// Команды по умолчанию
Command.stIo.xOpenDoor := FALSE;
Command.stIo.xCloseDoor := FALSE;
Command.stIo.xHatchUnLock := FALSE;
Command.stIo.xOpenSafetyDoor := FALSE;
Command.stIo.xCloseSafetyDoor := FALSE;
Command.stIo.xClampChuck := FALSE;
Command.stIo.xUnclampChuck := FALSE;
Command.stIo.xStartCycle := FALSE;
Command.stIo.xReset := xReset OR xResetGlobal;

Command.stRobot.xExecute := FALSE;
Command.stRobot.xStop := FALSE;

// Импульсы ручного управления проходят только через рассчитанные PLC-разрешения.
// Автоматический алгоритм станка в DISABLED не формирует параллельных команд.
IF xHmiOpenSafetyDoor AND xManualSafetyDoorOpenAllowed THEN
	Command.stIo.xOpenSafetyDoor := TRUE;
END_IF;
IF xHmiCloseSafetyDoor AND xManualSafetyDoorCloseAllowed THEN
	Command.stIo.xCloseSafetyDoor := TRUE;
END_IF;
IF xHmiOpenHatch AND xManualHatchOpenAllowed THEN
	xManualHatchOpenDemand := TRUE;
	xManualHatchUnlockDemand := TRUE;
END_IF;
IF xHmiCloseHatch AND xManualHatchCloseAllowed THEN
	Command.stIo.xCloseDoor := TRUE;
	xManualHatchOpenDemand := FALSE;
	xManualHatchUnlockDemand := FALSE;
END_IF;
IF rtHmiUnlockHatch.Q AND xManualHatchUnlockAllowed THEN
	xManualHatchUnlockDemand := TRUE;
END_IF;
IF rtHmiLockHatch.Q AND xManualHatchLockAllowed THEN
	xManualHatchUnlockDemand := FALSE;
	xManualHatchOpenDemand := FALSE;
END_IF;
IF NOT xManualMode THEN
	xManualHatchUnlockDemand := FALSE;
	xManualHatchOpenDemand := FALSE;
END_IF;
IF xHmiOpenChuck AND xManualChuckOpenAllowed THEN
	Command.stIo.xUnclampChuck := TRUE;
END_IF;
IF xHmiCloseChuck AND xManualChuckCloseAllowed THEN
	Command.stIo.xClampChuck := TRUE;
END_IF;
Command.stRobot.eAction := E_ROBOT_ACTION.NONE;
xServiceDoorOpenDemand := FALSE;
xServiceDoorCloseDemand := FALSE;
xServiceHatchUnlockDemand := FALSE;

IF xTestInitialize THEN
	Error.dwErrorActive := DWORD#0;
	Error.dwAlarmActive := DWORD#0;
	uiIndex := UINT#0;
	xDisableRequest := FALSE;
	xOperatorRunningCNC := FALSE;
	xOperatorClosingDoor := FALSE;
	xAutoCycleCommanded := FALSE;
	xCycleMeasureActive := FALSE;
	xCycleMeasureValid := FALSE;
	xRetreatStarted := FALSE;
	xRobotInsideMachine := FALSE;
	xFaultContextCaptured := FALSE;
	xRobotInsideAtFault := FALSE;
	xDoorRobotStopLatched := FALSE;
	xRobotStopRequired := FALSE;
	xRobotDone := FALSE;
	xServiceDoorCloseDemand := FALSE;
	xServiceDoorOpenDemand := FALSE;
	xServiceHatchUnlockDemand := FALSE;
	xManualHatchUnlockDemand := FALSE;
	xManualHatchOpenDemand := FALSE;
	xAutoDoorOpenLatched := FALSE;
	xRobotActionDone := FALSE;
	xRobotCommandStarted := FALSE;
	eGrantedOperation := E_MACHINE_OPERATION.NONE;
	eActualOperation := E_MACHINE_OPERATION.NONE;
	IF (uiTestInitialState = UINT#0) OR NOT xPointsConfigured THEN
		eState := E_MACHINE_STATE.DISABLED;
		ePartType := E_PART_TYPE.UNKNOWN;
	ELSE
		eState := E_MACHINE_STATE.IDLE;
		IF uiTestInitialState = UINT#3 THEN
			ePartType := E_PART_TYPE.DETAIL;
		ELSIF uiTestInitialState = UINT#2 THEN
			ePartType := E_PART_TYPE.PART;
		ELSE
			ePartType := E_PART_TYPE.UNKNOWN;
		END_IF;
	END_IF;
END_IF;

IF stMachineStatus.xChuckClamped AND NOT stMachineStatus.xAlarm THEN
	ePartState := E_PART_STATE.LOADED;
ELSIF stMachineStatus.xChuckUnclamped AND NOT stMachineStatus.xAlarm THEN
	ePartState := E_PART_STATE.EMPTY;
ELSE
	ePartState := E_PART_STATE.UNKNOWN;
END_IF


// // Ручное подтверждение состояния детали
// IF (eState = E_MACHINE_STATE.IDLE)
// AND NOT stMachineStatus.xCycleActive THEN
//     IF rtSetPartLoaded.Q THEN
//         ePartState := E_PART_STATE.LOADED;
//     END_IF;
// 
//     IF rtSetPartEmpty.Q THEN
//         ePartState := E_PART_STATE.EMPTY;
//     END_IF;
// END_IF;

// Автоматическое открытие после окончания обработки
IF rtCycleDone.Q 
	AND NOT stMachineStatus.xAlarm 
	AND NOT stMachineStatus.xCycleActive 
	AND (eState = E_MACHINE_STATE.IDLE) 
	AND NOT xGlobalError THEN
	ePartType := E_PART_TYPE.DETAIL;
    xAutoDoorOpenLatched := TRUE;
END_IF;

IF stMachineStatus.xDoorOpen THEN
    xAutoDoorOpenLatched := FALSE;
END_IF;

eGrantedOperation := E_MACHINE_OPERATION.NONE;

IF (ePartState = E_PART_STATE.EMPTY)
AND (ePartType = E_PART_TYPE.UNKNOWN)
AND stRobotStatus.xBlankAvailable  THEN
    eGrantedOperation := E_MACHINE_OPERATION.LOAD;

ELSIF (ePartState = E_PART_STATE.LOADED)
AND (ePartType = E_PART_TYPE.DETAIL) THEN
    IF stRobotStatus.xBlankAvailable THEN
        eGrantedOperation := E_MACHINE_OPERATION.CHANGE;
    ELSE
        eGrantedOperation := E_MACHINE_OPERATION.UNLOAD;
    END_IF;
ELSIF (ePartState = E_PART_STATE.UNKNOWN) THEN
	eGrantedOperation := E_MACHINE_OPERATION.NONE;
END_IF;

// Включение и отключение блока
IF xDisableRequest
AND ((eState = E_MACHINE_STATE.IDLE)
	OR (eState = E_MACHINE_STATE.OPERATOR_CHOICE_PART)
	OR (eState = E_MACHINE_STATE.OPERATOR_CHOICE_DOOR)
	OR (eState = E_MACHINE_STATE.OPERATOR_CHOICE_RUN)) THEN
    eState := E_MACHINE_STATE.DISABLED;
ELSIF rtEnabledMachine.Q
AND NOT rtDisabledMachine.Q
AND (eState = E_MACHINE_STATE.DISABLED) THEN
	IF NOT stMachineStatus.xAlarm
	AND NOT stMachineStatus.xCycleActive
	AND xSafetyDoorSafe
	AND xPointsConfigured THEN
		IF ePartState = E_PART_STATE.EMPTY THEN
			eState := E_MACHINE_STATE.IDLE;
		ELSIF ePartState = E_PART_STATE.LOADED THEN
			eState := E_MACHINE_STATE.OPERATOR_CHOICE_PART;
		END_IF;
	END_IF;
END_IF;

IF xGlobalError
AND (eState <> E_MACHINE_STATE.DISABLED) THEN
    Error.dwErrorActive := Error.dwErrorActive OR ERR_SAFETY_STOP;
    eState := E_MACHINE_STATE.ERROR;
END_IF;

IF stMachineStatus.xAlarm AND (eState = E_MACHINE_STATE.IDLE) THEN
	Error.dwErrorActive := Error.dwErrorActive OR ERR_MACHINE_IDLE;
    eState := E_MACHINE_STATE.ERROR;
END_IF

IF ((eState = E_MACHINE_STATE.OPERATOR_CHOICE_PART) OR (eState = E_MACHINE_STATE.OPERATOR_CHOICE_DOOR) OR (eState = E_MACHINE_STATE.OPERATOR_CHOICE_RUN))
AND ftChuckClamped.Q THEN
	eState := E_MACHINE_STATE.DISABLED;
END_IF; 

IF (eState = E_MACHINE_STATE.DISABLED) OR (eState = E_MACHINE_STATE.ERROR) THEN
	xOperatorRunningCNC := FALSE;
	xOperatorClosingDoor := FALSE;
	ePartType :=   E_PART_TYPE.UNKNOWN;
END_IF
// Останавливаем робота, если люк закрылся при нахождении робота в станке.
tofErrorDoor(
			PT:= T#100MS,
			IN:=stMachineStatus.xDoorOpen
);

// Ошибка робота в рабочей зоне принадлежит одновременно роботу и станку.
// Для действия захвата сохраняется отдельная диагностическая причина.
IF xRobotInsideMachine
AND stRobotStatus.xError
AND (eState <> E_MACHINE_STATE.ERROR) THEN
	IF eState = E_MACHINE_STATE.ROBOT_ACTION THEN
		Error.dwErrorActive := Error.dwErrorActive OR ERR_ROBOT_ACTION;
	ELSE
		Error.dwErrorActive := Error.dwErrorActive OR ERR_ROBOT_MOTION;
	END_IF;
	eState := E_MACHINE_STATE.ERROR;
END_IF;
						
IF xRobotInsideMachine
AND (
	(rtDoorClosed.Q)
	OR (
		NOT tofErrorDoor.Q
		AND (stRobotStatus.xBusy
			OR (eState = E_MACHINE_STATE.ROBOT_MOVE)
			OR (eState = E_MACHINE_STATE.ROBOT_ACTION))
	)
) THEN
	// Stop должен быть явным даже при гонке статусов: xBusy уже мог успеть
	// сброситься в FB_ROBOT, пока группа ещё принимает команду останова.
	Command.stRobot.xStop := TRUE;
	xDoorRobotStopLatched := TRUE;
	Error.dwErrorActive := Error.dwErrorActive OR ERR_DOOR_ROBOT;
    eState := E_MACHINE_STATE.ERROR;
END_IF

// Открытие операторской двери в любой момент роботного обслуживания
// — первичная авария станка с каскадным ROBOT_STOP.
IF (eActualOperation <> E_MACHINE_OPERATION.NONE)
AND NOT xManualMode
AND NOT xSafetyDoorSafe
AND (eState <> E_MACHINE_STATE.ERROR) THEN
	Command.stRobot.xStop := stRobotStatus.xBusy;
	Error.dwErrorActive := Error.dwErrorActive OR ERR_SAFETY_DOOR_OPEN;
	eState := E_MACHINE_STATE.ERROR;
END_IF;

// Старый рецепт и удерживаемые запросы не возобновляются после ручного I/O.
// Состояние патрона будет повторно определено при отдельном включении станка.
IF xIoManual THEN
	uiIndex := UINT#0;
	eActualOperation := E_MACHINE_OPERATION.NONE;
	eGrantedOperation := E_MACHINE_OPERATION.NONE;
	xRobotDone := FALSE;
	xRobotCommandStarted := FALSE;
	xManualHatchUnlockDemand := FALSE;
	xManualHatchOpenDemand := FALSE;
	xAutoDoorOpenLatched := FALSE;
	xOperatorRunningCNC := FALSE;
	xOperatorClosingDoor := FALSE;
	IF eState <> E_MACHINE_STATE.ERROR THEN
		eState := E_MACHINE_STATE.DISABLED;
	END_IF;
END_IF;

CASE eState OF
	E_MACHINE_STATE.DISABLED:
		xDisableRequest := FALSE;
		IF NOT stMachineStatus.xCycleActive THEN
			xAutoCycleCommanded := FALSE;
		END_IF;
		
	E_MACHINE_STATE.OPERATOR_CHOICE_PART:
		IF rtSetDetailLoaded.Q AND NOT stMachineStatus.xAlarm THEN
			eState := E_MACHINE_STATE.IDLE;
			ePartType := E_PART_TYPE.DETAIL;
		ELSIF rtSetBlankLoaded.Q AND NOT stMachineStatus.xAlarm THEN
			ePartType := E_PART_TYPE.PART;
			IF stMachineStatus.xDoorClosed THEN
				eState := E_MACHINE_STATE.OPERATOR_CHOICE_RUN;
			ELSE
				eState := E_MACHINE_STATE.OPERATOR_CHOICE_DOOR;
			END_IF;
		ELSIF stMachineStatus.xAlarm THEN
			Error.dwErrorActive := Error.dwErrorActive OR ERR_MACHINE_ALARM;
    		eState := E_MACHINE_STATE.ERROR;
		END_IF;
		
	E_MACHINE_STATE.OPERATOR_CHOICE_DOOR:
		// При уже закрытой двери шаг подтверждения закрытия не нужен:
		// автомат сразу переходит к вопросу о запуске обработки.
		IF stMachineStatus.xAlarm THEN
			Error.dwErrorActive := Error.dwErrorActive OR ERR_MACHINE_ALARM;
    		eState := E_MACHINE_STATE.ERROR;
		ELSIF xHmiRejectDoor THEN
			eState := E_MACHINE_STATE.DISABLED;
		ELSIF stMachineStatus.xDoorClosed THEN
			eState := E_MACHINE_STATE.OPERATOR_CHOICE_RUN;
		ELSIF xHmiAcceptDoor THEN
			xOperatorClosingDoor := TRUE;
			eState := E_MACHINE_STATE.DOOR_CLOSE;
		END_IF;
		
	E_MACHINE_STATE.OPERATOR_CHOICE_RUN:
		IF xHmiAcceptRunCNC AND NOT stMachineStatus.xAlarm THEN
			xOperatorRunningCNC := TRUE; 
			eState := E_MACHINE_STATE.CYCLE_START;
		ELSIF xHmiRejectRunCNC AND NOT stMachineStatus.xAlarm THEN
			eState := E_MACHINE_STATE.DISABLED;
		ELSIF stMachineStatus.xAlarm THEN
			Error.dwErrorActive := Error.dwErrorActive OR ERR_MACHINE_ALARM;
    		eState := E_MACHINE_STATE.ERROR;
		END_IF; 	
		
	E_MACHINE_STATE.IDLE:
		uiIndex := 0;
		xRobotDone := FALSE;
		IF xExecute THEN
			IF (stRobotStatus.eCurrentPoint = stPoints.eAbove)
			AND ePartState <> E_PART_STATE.UNKNOWN
			AND NOT stMachineStatus.xAlarm
			AND NOT stMachineStatus.xCycleActive
			AND xSafetyDoorSafe
    		AND NOT stRobotStatus.xBusy 
			AND NOT stRobotStatus.xError
			AND NOT xGlobalError THEN
				eActualOperation := eGrantedOperation;
				eState := E_MACHINE_STATE.CHOSE;
			ELSIF ePartState = E_PART_STATE.UNKNOWN THEN
				Error.dwErrorActive := Error.dwErrorActive OR ERR_UNKNOWN_DETAIL;
				eState := E_MACHINE_STATE.ERROR ;
			END_IF
		END_IF
		
	E_MACHINE_STATE.CHOSE:
		CASE eActualOperation OF 
			E_MACHINE_OPERATION.CHANGE:
				stRecipe := stChangeRecipe;
				eState := E_MACHINE_STATE.READ;
			E_MACHINE_OPERATION.LOAD:
				stRecipe := stLoadRecipe;
				eState := E_MACHINE_STATE.READ;
			E_MACHINE_OPERATION.UNLOAD:
				stRecipe := stUnloadRecipe;
				eState := E_MACHINE_STATE.READ;
		ELSE
			Error.dwErrorActive := Error.dwErrorActive OR ERR_WRONG_OPERATION ;
			eState := E_MACHINE_STATE.ERROR;
		END_CASE
		
	E_MACHINE_STATE.READ:
		CASE stRecipe[uiIndex].eCommand OF
			E_MACHINE_STATE.ROBOT_MOVE:
				xRobotCommandStarted := FALSE;
				eState := E_MACHINE_STATE.ROBOT_MOVE;
				
			E_MACHINE_STATE.ROBOT_ACTION:
				xRobotCommandStarted := FALSE;
				eState := E_MACHINE_STATE.ROBOT_ACTION;
				
			E_MACHINE_STATE.DOOR_OPEN:
				eState := E_MACHINE_STATE.DOOR_OPEN;
				
			E_MACHINE_STATE.DOOR_CLOSE:
				eState := E_MACHINE_STATE.DOOR_CLOSE;
				
			E_MACHINE_STATE.CHUCK_OPEN:
				eState := E_MACHINE_STATE.CHUCK_OPEN;
				
			E_MACHINE_STATE.CHUCK_CLOSE:
				eState := E_MACHINE_STATE.CHUCK_CLOSE;
				
			E_MACHINE_STATE.CYCLE_START:
				eState := E_MACHINE_STATE.CYCLE_START;
				
			E_MACHINE_STATE.DONE:
				eState := E_MACHINE_STATE.DONE;
				
		ELSE
			Error.dwErrorActive := Error.dwErrorActive OR ERR_WRONG_COMMAND;
			eState := E_MACHINE_STATE.ERROR;
		END_CASE
	
	E_MACHINE_STATE.NEXT:
			uiIndex := uiIndex + 1;
			IF uiIndex > 40 THEN
				Error.dwErrorActive := Error.dwErrorActive OR ERR_INDEX;
				eState := E_MACHINE_STATE.ERROR;
			ELSE
				eState := E_MACHINE_STATE.READ;
			END_IF;
	
	E_MACHINE_STATE.ROBOT_MOVE:
		Command.stRobot.xExecute  := TRUE;
		Command.stRobot.eAction   := E_ROBOT_ACTION.MOVE_TO_POINT;
		xRetreatStarted          := stRecipe[uiIndex].xRetreatStarted;
		IF stRecipe[uiIndex].stPoint = E_MACHINE_POINTS.ABOVE  THEN
			Command.stRobot.eSetPoint := stPoints.eAbove;
		ELSIF stRecipe[uiIndex].stPoint = E_MACHINE_POINTS.CHUCK THEN
			Command.stRobot.eSetPoint := stPoints.eChuck;
		ELSIF stRecipe[uiIndex].stPoint = E_MACHINE_POINTS.CHUCK_APPROACH THEN
			Command.stRobot.eSetPoint := stPoints.eChuckApproach;
		ELSIF stRecipe[uiIndex].stPoint = E_MACHINE_POINTS.INSIDE THEN
			Command.stRobot.eSetPoint := stPoints.eInside;
		END_IF
		IF stRobotStatus.xBusy THEN
			xRobotCommandStarted := TRUE;
		END_IF;

		IF stRobotStatus.xError THEN
			Error.dwErrorActive := Error.dwErrorActive OR ERR_ROBOT_MOTION;
			eState := E_MACHINE_STATE.ERROR ;
			
		ELSIF stMachineStatus.xAlarm THEN
			Command.stRobot.xStop := stRobotStatus.xBusy;
			Error.dwErrorActive := Error.dwErrorActive OR ERR_MACHINE_ALARM;
			eState := E_MACHINE_STATE.ERROR ;
			
		ELSIF xRobotCommandStarted AND stRobotStatus.xDone THEN
        	eState := E_MACHINE_STATE.RELEASE_ROBOT_ACTION;

		ELSIF tonRobotMoveTimeout.Q THEN
			Command.stRobot.xStop := stRobotStatus.xBusy;
			Error.dwErrorActive := Error.dwErrorActive OR ERR_TIMEOUT_ROBOT_MOVE;
			eState := E_MACHINE_STATE.ERROR;
			
    	END_IF;
	
	E_MACHINE_STATE.ROBOT_ACTION:
		xRobotActionDone := FALSE;

		CASE stRecipe[uiIndex].eRobotAction OF
			E_ROBOT_ACTION.UNCLAMP_1:
				xRobotActionDone := stRobotStatus.xGripper1Open;
			E_ROBOT_ACTION.CLAMP_1:
				xRobotActionDone := stRobotStatus.xGripper1Closed;
			E_ROBOT_ACTION.UNCLAMP_2:
				xRobotActionDone := stRobotStatus.xGripper2Open;
			E_ROBOT_ACTION.CLAMP_2:
				xRobotActionDone := stRobotStatus.xGripper2Closed;
			E_ROBOT_ACTION.ROTATE_TO_BLANK:
				xRobotActionDone := stRobotStatus.xRotatedToBlank;
			E_ROBOT_ACTION.ROTATE_TO_DETAIL:
				xRobotActionDone := stRobotStatus.xRotatedToDetail;
		END_CASE;
		IF xRobotActionDone THEN
			eState := E_MACHINE_STATE.NEXT;
		ELSE
			Command.stRobot.xExecute := TRUE;
			Command.stRobot.eAction := stRecipe[uiIndex].eRobotAction;
		END_IF;
		IF stRobotStatus.xBusy THEN
			xRobotCommandStarted := TRUE;
		END_IF;
		
		IF (eState = E_MACHINE_STATE.ROBOT_ACTION)
		AND stMachineStatus.xAlarm THEN
			Command.stRobot.xStop := stRobotStatus.xBusy;
			Error.dwErrorActive := Error.dwErrorActive OR ERR_MACHINE_ALARM;
			eState := E_MACHINE_STATE.ERROR ;
	
		ELSIF (eState = E_MACHINE_STATE.ROBOT_ACTION)
		AND stRobotStatus.xError THEN
			Error.dwErrorActive := Error.dwErrorActive OR ERR_ROBOT_ACTION;
			eState := E_MACHINE_STATE.ERROR ;

		ELSIF (eState = E_MACHINE_STATE.ROBOT_ACTION)
		AND tonRobotActionTimeout.Q THEN
			Command.stRobot.xStop := stRobotStatus.xBusy;
			Error.dwErrorActive := Error.dwErrorActive OR ERR_TIMEOUT_ROBOT_ACTION;
			eState := E_MACHINE_STATE.ERROR;
			
		ELSIF (eState = E_MACHINE_STATE.ROBOT_ACTION)
		AND xRobotCommandStarted
		AND stRobotStatus.xDone THEN
        	eState := E_MACHINE_STATE.RELEASE_ROBOT_ACTION;
    	END_IF;
		
	E_MACHINE_STATE.RELEASE_ROBOT_ACTION:
		IF NOT stRobotStatus.xBusy
    	AND NOT stRobotStatus.xDone
		AND NOT stRobotStatus.xError THEN
			xRobotDone := stRecipe[uiIndex].xRobotDone;
        	eState := E_MACHINE_STATE.NEXT;
			
		ELSIF stRobotStatus.xError AND  stRecipe[uiIndex].eRobotAction = E_ROBOT_ACTION.MOVE_TO_POINT THEN
			Error.dwErrorActive := Error.dwErrorActive OR ERR_ROBOT_MOTION;
			eState := E_MACHINE_STATE.ERROR;
			
		ELSIF stRobotStatus.xError THEN
			Error.dwErrorActive := Error.dwErrorActive OR ERR_ROBOT_ACTION;
			eState := E_MACHINE_STATE.ERROR;

		ELSIF tonRobotReleaseTimeout.Q THEN
			Command.stRobot.xStop := stRobotStatus.xBusy;
			Error.dwErrorActive := Error.dwErrorActive OR ERR_TIMEOUT_ROBOT_RELEASE;
			eState := E_MACHINE_STATE.ERROR;
    	END_IF;
		
	E_MACHINE_STATE.DOOR_OPEN:
		xServiceDoorOpenDemand := TRUE;
		// Сначала снимаем замок, затем открываем роботный люк.
		IF stMachineStatus.xHatchLocked THEN
			xServiceHatchUnlockDemand := TRUE;
		END_IF;

	    IF stMachineStatus.xDoorOpen
		AND NOT stMachineStatus.xHatchLocked
		AND NOT stMachineStatus.xAlarm THEN
			xServiceDoorOpenDemand := FALSE;
			xServiceHatchUnlockDemand := FALSE;
         	eState := E_MACHINE_STATE.NEXT;
		ELSIF stMachineStatus.xAlarm THEN
			Error.dwErrorActive := Error.dwErrorActive OR ERR_DOOR_OPEN;
			eState := E_MACHINE_STATE.ERROR;
		ELSIF tonDoorOpenTimeout.Q THEN
			xServiceDoorOpenDemand := FALSE;
			Error.dwErrorActive := Error.dwErrorActive OR ERR_TIMEOUT_DOOR_OPEN;
			eState := E_MACHINE_STATE.ERROR;
    	END_IF;
	
	E_MACHINE_STATE.DOOR_CLOSE: 
		// После сервисной операции безопасность подтверждает защёлка xRobotDone:
		// рецепт уже довёл робот до ABOVE и освободил его для следующего маршрута.
		// Общий xBusy больше не блокирует дверь: робот может двигаться к другому узлу.
		IF xRobotInsideMachine
		OR (NOT xOperatorClosingDoor AND NOT xRobotDone) THEN
			Command.stRobot.xStop := xRobotInsideMachine AND stRobotStatus.xBusy;
			xDoorRobotStopLatched := TRUE;
			Error.dwErrorActive := Error.dwErrorActive OR ERR_DOOR_ROBOT;
			eState := E_MACHINE_STATE.ERROR;
		ELSE
			xServiceDoorCloseDemand := TRUE;
			// Замок удерживается открытым до подтверждения закрытой двери.
			IF NOT stMachineStatus.xDoorClosed THEN
				xServiceHatchUnlockDemand := TRUE;
			END_IF;
		END_IF;

		IF stMachineStatus.xDoorClosed THEN
			xServiceHatchUnlockDemand := FALSE;
		END_IF;
		IF (eState = E_MACHINE_STATE.DOOR_CLOSE)
		AND stMachineStatus.xDoorClosed
		AND stMachineStatus.xHatchLocked
		AND NOT stMachineStatus.xAlarm THEN
			xServiceDoorCloseDemand := FALSE;
			IF NOT xOperatorClosingDoor THEN
				eState := E_MACHINE_STATE.NEXT;
			ELSIF xOperatorClosingDoor THEN
				eState := E_MACHINE_STATE.OPERATOR_CHOICE_RUN;
				xOperatorClosingDoor := FALSE;
			END_IF;
		ELSIF stMachineStatus.xAlarm THEN
			Error.dwErrorActive := Error.dwErrorActive OR ERR_DOOR_CLOSE;
			eState := E_MACHINE_STATE.ERROR;
		ELSIF (eState = E_MACHINE_STATE.DOOR_CLOSE)
		AND tonDoorCloseTimeout.Q THEN
			xServiceDoorCloseDemand := FALSE;
			Error.dwErrorActive := Error.dwErrorActive OR ERR_TIMEOUT_DOOR_CLOSE;
			eState := E_MACHINE_STATE.ERROR;
    	END_IF;
		
	E_MACHINE_STATE.CHUCK_OPEN: 
		Command.stIo.xUnclampChuck := TRUE;

    	IF stMachineStatus.xChuckUnclamped 
		AND NOT stMachineStatus.xAlarm THEN
			Command.stIo.xUnclampChuck := FALSE;
			ePartType := E_PART_TYPE.UNKNOWN;
       		eState := E_MACHINE_STATE.NEXT;
		ELSIF stMachineStatus.xAlarm THEN
			Command.stIo.xUnclampChuck := FALSE;
			Error.dwErrorActive := Error.dwErrorActive OR ERR_CHUCK_OPEN;
			eState := E_MACHINE_STATE.ERROR;
		ELSIF tonChuckOpenTimeout.Q THEN
			Command.stIo.xUnclampChuck := FALSE;
			Error.dwErrorActive := Error.dwErrorActive OR ERR_TIMEOUT_CHUCK_OPEN;
			eState := E_MACHINE_STATE.ERROR;
    	END_IF;
		
	
	E_MACHINE_STATE.CHUCK_CLOSE: 
		Command.stIo.xClampChuck := TRUE;

    	IF stMachineStatus.xChuckClamped 
		AND NOT stMachineStatus.xAlarm THEN
			Command.stIo.xClampChuck := FALSE;
			ePartType := E_PART_TYPE.PART;
       		eState := E_MACHINE_STATE.NEXT;
		ELSIF stMachineStatus.xAlarm THEN
			Command.stIo.xClampChuck := FALSE;
			Error.dwErrorActive := Error.dwErrorActive OR ERR_CHUCK_CLOSE;
			eState := E_MACHINE_STATE.ERROR;
		ELSIF tonChuckCloseTimeout.Q THEN
			Command.stIo.xClampChuck := FALSE;
			Error.dwErrorActive := Error.dwErrorActive OR ERR_TIMEOUT_CHUCK_CLOSE;
			eState := E_MACHINE_STATE.ERROR;
    	END_IF;
		
	E_MACHINE_STATE.CYCLE_START:
		IF stMachineStatus.xChuckClamped
    	AND stMachineStatus.xDoorClosed THEN
			Command.stIo.xStartCycle := TRUE;
			xAutoCycleCommanded := TRUE;
		END_IF;
		
        IF stMachineStatus.xCycleActive
		AND NOT stMachineStatus.xAlarm THEN
			Command.stIo.xStartCycle := FALSE;
			IF NOT xOperatorRunningCNC THEN
            	eState := E_MACHINE_STATE.NEXT;
			ELSIF xOperatorRunningCNC THEN
				xOperatorRunningCNC := FALSE;
				eState := E_MACHINE_STATE.IDLE;
			END_IF;
		ELSIF stMachineStatus.xAlarm THEN
			Command.stIo.xStartCycle := FALSE;
			Error.dwErrorActive := Error.dwErrorActive OR ERR_CYCLE_START;
			eState := E_MACHINE_STATE.ERROR;
		ELSIF tonCycleStartTimeout.Q THEN
			Command.stIo.xStartCycle := FALSE;
			xAutoCycleCommanded := FALSE;
			Error.dwErrorActive := Error.dwErrorActive OR ERR_TIMEOUT_CYCLE_START;
			eState := E_MACHINE_STATE.ERROR;
        END_IF;
	
	E_MACHINE_STATE.DONE:
		CASE eActualOperation OF 
			E_MACHINE_OPERATION.CHANGE, E_MACHINE_OPERATION.LOAD:
				eActualOperation := E_MACHINE_OPERATION.NONE;
				ePartState := E_PART_STATE.LOADED;						
			E_MACHINE_OPERATION.UNLOAD:
				eActualOperation := E_MACHINE_OPERATION.NONE;
				ePartState := E_PART_STATE.EMPTY;
		END_CASE
		
		IF NOT xExecute THEN
			xRobotDone := FALSE;	
			eState := E_MACHINE_STATE.IDLE;
		END_IF
		
    E_MACHINE_STATE.ERROR:
		uiIndex := 0;
		eActualOperation := E_MACHINE_OPERATION.NONE;
		eGrantedOperation := E_MACHINE_OPERATION.NONE;
		IF NOT stMachineStatus.xCycleActive THEN
			xAutoCycleCommanded := FALSE;
		END_IF;

		IF (xReset OR xResetGlobal)
		AND NOT xIoManual
		AND NOT xGlobalError
		AND NOT xExecute
		AND NOT stMachineStatus.xAlarm
		AND xSafetyDoorSafe
		AND xDoorRobotRecoveryReady
		AND xRobotResetDependencyReady THEN
			Error.dwErrorLast := Error.dwErrorActive;
			Error.dwErrorActive := DWORD#0;
			xManualHatchUnlockDemand := FALSE;
			xManualHatchOpenDemand := FALSE;
        	eState := E_MACHINE_STATE.DISABLED;
    	END_IF;
END_CASE;

// Таймаут одинаково контролирует автоматическое и ручное снятие замка.
// После отказа удерживаемый запрос снимается, чтобы сброс не запустил его
// повторно без нового явного действия оператора.
IF tonHatchUnlockTimeout.Q
AND (eState <> E_MACHINE_STATE.ERROR) THEN
	xServiceHatchUnlockDemand := FALSE;
	xManualHatchUnlockDemand := FALSE;
	xManualHatchOpenDemand := FALSE;
	Error.dwErrorActive := Error.dwErrorActive OR ERR_TIMEOUT_HATCH_UNLOCK;
	eState := E_MACHINE_STATE.ERROR;
END_IF;

// Причина остаётся в своём CASE, а единая реакция рассчитывается один раз.
// Контекст защёлкивается до сброса, поэтому смена состояния робота его не теряет.
IF (eState = E_MACHINE_STATE.ERROR) AND NOT xFaultContextCaptured THEN
	xRobotInsideAtFault := xRobotInsideMachine;
	xFaultContextCaptured := TRUE;
ELSIF eState <> E_MACHINE_STATE.ERROR THEN
	xRobotInsideAtFault := FALSE;
	xFaultContextCaptured := FALSE;
END_IF;

xRobotStopRequired := NOT xGlobalError
	AND (
		((Error.dwErrorActive
			AND (MASK_ALWAYS_ROBOT_STOP AND NOT ERR_DOOR_ROBOT)) <> DWORD#0)
		OR (((Error.dwErrorActive AND ERR_DOOR_ROBOT) <> DWORD#0)
			AND NOT xDoorRobotRecoveryReady)
		OR xDoorRobotStopLatched
		OR (((Error.dwErrorActive
			AND (MASK_EQUIPMENT_ERROR AND NOT ERR_DOOR_ROBOT)) <> DWORD#0)
			AND xRobotInsideAtFault)
	);

// Stop нужен только выполняемому действию. Стоящий в станке робот получает
// зависимую ошибку через FB_ROBOT, но бессмысленная команда Stop не выдаётся.
IF (eState = E_MACHINE_STATE.ERROR)
AND xRobotStopRequired
AND (stRobotStatus.xBusy OR xRobotMotionBusy) THEN
	Command.stRobot.xStop := TRUE;
END_IF;

// После подтверждённого открытия люка и полной остановки можно отпустить
// защёлку зависимого Stop; до этого новый цикл не должен стартовать.
IF xDoorRobotStopLatched
AND NOT xRobotMotionBusy
AND xDoorRobotRecoveryReady THEN
	xDoorRobotStopLatched := FALSE;
END_IF;

IF ((eState <> E_MACHINE_STATE.ERROR) OR xManualHatchRecoveryOpenAllowed)
AND NOT xGlobalError AND NOT xIoManual THEN
	Command.stIo.xHatchUnLock := xManualHatchUnlockDemand OR xServiceHatchUnlockDemand;
	IF xManualHatchOpenDemand
	AND NOT stMachineStatus.xHatchLocked
	AND NOT stMachineStatus.xDoorOpen
	AND NOT stMachineStatus.xCycleActive
	AND NOT stMachineStatus.xAlarm THEN
		Command.stIo.xOpenDoor := TRUE;
	END_IF;
    IF (eState <> E_MACHINE_STATE.ERROR) AND xServiceDoorCloseDemand 
	AND NOT (xAutoDoorOpenLatched OR xServiceDoorOpenDemand)
	AND NOT xRobotInsideMachine
	AND (xOperatorClosingDoor OR xRobotDone)
	AND NOT stMachineStatus.xAlarm THEN
        Command.stIo.xCloseDoor := TRUE;

    ELSIF (eState <> E_MACHINE_STATE.ERROR) AND (xAutoDoorOpenLatched OR xServiceDoorOpenDemand)
	AND NOT xServiceDoorCloseDemand
	AND NOT stMachineStatus.xHatchLocked
    AND NOT stMachineStatus.xCycleActive
    AND NOT stMachineStatus.xAlarm THEN
        Command.stIo.xOpenDoor := TRUE;
    END_IF;
END_IF;

// Замок нельзя открывать во время обработки выбранного для автоматической
// линии станка. Срабатывание формируется самим PLC по фактической команде.
IF xAutomaticUseEnabled
AND stMachineStatus.xCycleActive
AND NOT stMachineStatus.xHatchLocked THEN
	Command.stIo.xHatchUnLock := FALSE;
	Error.dwErrorActive := Error.dwErrorActive OR ERR_HATCH_UNLOCK_PROCESSING;
	eState := E_MACHINE_STATE.ERROR;
END_IF;

Status.xCanAcceptService := (eState = E_MACHINE_STATE.IDLE)
			AND ePartState <> E_PART_STATE.UNKNOWN
			AND NOT stMachineStatus.xAlarm
			AND NOT stMachineStatus.xCycleActive
			AND xSafetyDoorSafe
			AND NOT xGlobalError;

// В состоянии ERROR станок уже остановлен и не считается включённым.
// Это позволяет HMI показать команду «Включить станок», но оставить её
// недоступной до устранения причины и сброса ошибки.
Status.xEnabled := (eState <> E_MACHINE_STATE.DISABLED)
	AND (eState <> E_MACHINE_STATE.ERROR);
Status.xDisablePending := xDisableRequest AND Status.xEnabled;
Status.xPowerAllowed := (eState <> E_MACHINE_STATE.ERROR)
	AND (xDisableRequest
		OR (eState <> E_MACHINE_STATE.DISABLED)
		OR ((eState = E_MACHINE_STATE.DISABLED)
			AND xPointsConfigured
			AND NOT stMachineStatus.xAlarm
			AND NOT stMachineStatus.xCycleActive
			AND xSafetyDoorSafe
			AND (ePartState <> E_PART_STATE.UNKNOWN)));
Status.xResetAllowed := (eState = E_MACHINE_STATE.ERROR)
	AND NOT xIoManual
	AND (Error.dwErrorActive <> DWORD#0)
	AND NOT stMachineStatus.xAlarm
	AND xSafetyDoorSafe
	AND NOT xGlobalError
	AND NOT xExecute
	AND (((Error.dwErrorActive AND ERR_DOOR_ROBOT) = DWORD#0)
		OR xDoorRobotRecoveryReady)
	AND xRobotResetDependencyReady;
Status.xManualControlAllowed := xManualControlAllowed;
Status.xManualSafetyDoorControlEnabled := xSafetyDoorControlEnabled;
Status.xManualSafetyDoorOpenAllowed := xManualSafetyDoorOpenAllowed;
Status.xManualSafetyDoorCloseAllowed := xManualSafetyDoorCloseAllowed;
Status.xManualHatchOpenAllowed := xManualHatchOpenAllowed;
Status.xManualHatchCloseAllowed := xManualHatchCloseAllowed;
Status.xManualHatchUnlockAllowed := xManualHatchUnlockAllowed;
Status.xManualHatchLockAllowed := xManualHatchLockAllowed;
Status.xManualChuckOpenAllowed := xManualChuckOpenAllowed;
Status.xManualChuckCloseAllowed := xManualChuckCloseAllowed;
Status.xProcessing := stMachineStatus.xCycleActive;
Status.xPartReady := stMachineStatus.xCycleDone;
Status.xServiceRequired := (eGrantedOperation <> E_MACHINE_OPERATION.NONE)
	AND (eState = E_MACHINE_STATE.IDLE);
Status.xRobotReleased := xRobotDone;
Status.xDone := (eState = E_MACHINE_STATE.DONE);
Status.xBusy :=  (eState <> E_MACHINE_STATE.IDLE)
				AND (eState <> E_MACHINE_STATE.DISABLED)
				AND (eState <> E_MACHINE_STATE.ERROR)
				AND (eState <> E_MACHINE_STATE.DONE)
				AND (eState <> E_MACHINE_STATE.OPERATOR_CHOICE_PART)
				AND (eState <> E_MACHINE_STATE.OPERATOR_CHOICE_RUN)
				AND (eState <> E_MACHINE_STATE.OPERATOR_CHOICE_DOOR)
				AND NOT ((eState = E_MACHINE_STATE.CYCLE_START) AND xOperatorRunningCNC)
				AND NOT ((eState = E_MACHINE_STATE.DOOR_CLOSE) AND xOperatorClosingDoor);
Status.xError := (eState = E_MACHINE_STATE.ERROR);
Status.xCriticalError := xRobotStopRequired;
Status.xAlarmError    := (Error.dwErrorActive AND MASK_EQUIPMENT_ERROR) <> DWORD#0;
Status.xExternalError := (Error.dwErrorActive AND MASK_EXTERNAL_ERROR) <> DWORD#0;
Status.xServiceRejected := (Error.dwErrorActive
	AND (ERR_DOOR_OPEN OR ERR_TIMEOUT_DOOR_OPEN)) <> DWORD#0
	AND ((Error.dwErrorActive
		AND NOT (ERR_DOOR_OPEN OR ERR_TIMEOUT_DOOR_OPEN)) = DWORD#0);
Error.dwAlarmActive := Error.dwErrorActive;
Status.xDoorOpen := stMachineStatus.xDoorOpen;
Status.xAlarm := stMachineStatus.xAlarm;
Status.eRecommendedOperation := eGrantedOperation;
Status.ePartState := ePartState;
Status.ePartType := ePartType;
Status.eAbovePoint := stPoints.eAbove;
Status.tCycleExpected := tExpectedCycle;
Status.tCycleElapsed := tonCycleMeasure.ET;
Status.tMeasuredCycle := tMeasuredCycle;
Status.xCycleTimeValid := tExpectedCycle > T#0S;
Status.xMeasuredTimeValid := xMeasuredTimeValid;
Status.xCycleOvertime := FALSE;
Status.tRemaining := T#0S;

IF stMachineStatus.xCycleActive
AND Status.xCycleTimeValid THEN
	IF Status.tCycleElapsed < Status.tCycleExpected THEN
		Status.tRemaining := Status.tCycleExpected - Status.tCycleElapsed;
	ELSE
		Status.xCycleOvertime := TRUE;
	END_IF;
END_IF;

Diag.eState := eState;
Diag.eGrantedOperation := eGrantedOperation;
Diag.eActualOperation := eActualOperation;

IF Error.dwErrorActive <> DWORD#0 THEN
	Error.dwErrorLast := Error.dwErrorActive;
END_IF;

Error.stErrorActive := UpdateErrorView(dwError := Error.dwErrorActive);
Error.stErrorLast := UpdateErrorView(dwError := Error.dwErrorLast);

METHOD UpdateErrorView : ST_MACHINE_ERROR
VAR_INPUT
	dwError : DWORD; // Битовая маска для расшифровки
END_VAR
VAR
	stError : ST_MACHINE_ERROR; // Представление ошибок отдельными флагами
END_VAR
stError.WRONG_OPERATION := (dwError AND ERR_WRONG_OPERATION) <> DWORD#0;
stError.WRONG_COMMAND := (dwError AND ERR_WRONG_COMMAND) <> DWORD#0;
stError.ROBOT_MOTION := (dwError AND ERR_ROBOT_MOTION) <> DWORD#0;
stError.ROBOT_ACTION := (dwError AND ERR_ROBOT_ACTION) <> DWORD#0;
stError.DOOR_OPEN := (dwError AND ERR_DOOR_OPEN) <> DWORD#0;
stError.DOOR_CLOSE := (dwError AND ERR_DOOR_CLOSE) <> DWORD#0;
stError.CHUCK_OPEN := (dwError AND ERR_CHUCK_OPEN) <> DWORD#0;
stError.CHUCK_CLOSE := (dwError AND ERR_CHUCK_CLOSE) <> DWORD#0;
stError.CYCLE_START := (dwError AND ERR_CYCLE_START) <> DWORD#0;
stError.SAFETY_STOP := (dwError AND ERR_SAFETY_STOP) <> DWORD#0;
stError.UNKNOWN_DETAIL := (dwError AND ERR_UNKNOWN_DETAIL) <> DWORD#0;
stError.MACHINE_ALARM := (dwError AND ERR_MACHINE_ALARM) <> DWORD#0;
stError.INDEX_ERROR := (dwError AND ERR_INDEX) <> DWORD#0;
stError.DOOR_ROBOT := (dwError AND ERR_DOOR_ROBOT) <> DWORD#0;
stError.MACHINE_IDLE := (dwError AND ERR_MACHINE_IDLE) <> DWORD#0;
stError.TIMEOUT_ROBOT_MOVE := (dwError AND ERR_TIMEOUT_ROBOT_MOVE) <> DWORD#0;
stError.TIMEOUT_ROBOT_ACTION := (dwError AND ERR_TIMEOUT_ROBOT_ACTION) <> DWORD#0;
stError.TIMEOUT_ROBOT_RELEASE := (dwError AND ERR_TIMEOUT_ROBOT_RELEASE) <> DWORD#0;
stError.TIMEOUT_DOOR_OPEN := (dwError AND ERR_TIMEOUT_DOOR_OPEN) <> DWORD#0;
stError.TIMEOUT_DOOR_CLOSE := (dwError AND ERR_TIMEOUT_DOOR_CLOSE) <> DWORD#0;
stError.TIMEOUT_HATCH_UNLOCK := (dwError AND ERR_TIMEOUT_HATCH_UNLOCK) <> DWORD#0;
stError.TIMEOUT_CHUCK_OPEN := (dwError AND ERR_TIMEOUT_CHUCK_OPEN) <> DWORD#0;
stError.TIMEOUT_CHUCK_CLOSE := (dwError AND ERR_TIMEOUT_CHUCK_CLOSE) <> DWORD#0;
stError.TIMEOUT_CYCLE_START := (dwError AND ERR_TIMEOUT_CYCLE_START) <> DWORD#0;
stError.SAFETY_DOOR_OPEN := (dwError AND ERR_SAFETY_DOOR_OPEN) <> DWORD#0;
stError.HATCH_UNLOCK_PROCESSING := (dwError AND ERR_HATCH_UNLOCK_PROCESSING) <> DWORD#0;

UpdateErrorView := stError;
END_METHOD

END_FUNCTION_BLOCK

// Device/Application/FB/FB_ROBOT
FUNCTION_BLOCK FB_ROBOT
VAR_INPUT
	xUsePhysicalGripperFeedback : BOOL;
	xPhysicalGripperIoReady : BOOL;
	stPhysicalGripperFeedback : ST_GRIPPER_STATUS;
	tPhysicalGripperActionTimeout : TIME := T#10S;
	axMagazineExchangeInProgress : ARRAY [1..2] OF BOOL; // Блокировка адресуется только к меняемому магазину
	xTestInitialize : BOOL;
	auiTestGripperContent : ARRAY [1..2] OF UINT;
	auiTestGripperType : ARRAY [1..2] OF UINT;
	uiTestOrientation : UINT;
	xExternalCommandInhibit : BOOL; // Программный экстренный останов запрещает следующую внешнюю команду
	xSimulationAccelerationEnable : BOOL; // Разрешить ускорение виртуальных таймеров только в симуляции
	uiSimulationTimeFactor : UINT := 1; // Коэффициент виртуального времени 1..100

	stMachine_1_Command : ST_ROBOT_COMMAND; // Команда роботу от первого станка
	stMachine_2_Command : ST_ROBOT_COMMAND; // Команда роботу от второго станка
	stMachine_3_Command : ST_ROBOT_COMMAND; // Команда роботу от третьего станка
	stMagazineCommand   : ST_ROBOT_COMMAND; // Команда роботу от магазина
	stCellCommand       : ST_ROBOT_COMMAND; // Команда позиционирования от менеджера ячейки
	uiBlankPayloadType  : UINT; // Тип заготовки из состояния цикла
	uiDetailPayloadType : UINT; // Тип готовой детали из состояния цикла
	stHmiCommand        : ST_ROBOT_COMMAND; // Ручная команда роботу с HMI
	xReset              : BOOL; // Сброс ошибок робота
    xMode               : BOOL; // Режим робота: TRUE — Modbus, FALSE — SoftMotion
	xManual      		: BOOL; // 1 - ручной режим работы, 0 - автоматический режим работы
	xGlobalError        : BOOL; // Глобальная ошибка ячейки
	xEquipmentStopRequired : BOOL; // Владелец оборудования требует зависимую ошибку робота
	xModbusBusy         : BOOL; // Внешний робот выполняет команду
	xModbusDone         : BOOL; // Внешний робот завершил команду
	xModbusError        : BOOL; // Ошибка обмена или внешнего робота
	stModbusStatus      : ST_ROBOT_MODBUS_STATUS; // Декодированная обратная связь SC-500
	xHmiDrivesEnable    : BOOL; // Исходный запрос HMI на включение приводов
	xHmiDrivesDisable   : BOOL; // Исходный запрос HMI на отключение приводов
	xHmiStop            : BOOL; // Исходный запрос HMI на остановку
	xHmiDrivesEnableAccepted : BOOL; // RunMotion принял запрос включения в исходном состоянии цикла
	xHmiDrivesDisableAccepted : BOOL; // RunMotion принял запрос отключения в исходном состоянии цикла
	xHmiStopAccepted    : BOOL; // RunMotion принял запрос остановки в исходном состоянии цикла
	xHmiDrivesEnableAllowed : BOOL; // Текущее разрешение включения от владельца Motion-слоя
	xHmiDrivesDisableAllowed : BOOL; // Текущее разрешение отключения от владельца Motion-слоя
	xHmiStopAllowed     : BOOL; // Текущее разрешение остановки от владельца Motion-слоя
	xHmiPermit          : BOOL; // Ручные команды HMI разрешены режимом ячейки
	xManualRecoveryAllowed : BOOL; // Разрешить включение приводов в аварийном ручном восстановлении
	xDrivesPowered      : BOOL; // Все три привода включены
	xDrivesOff          : BOOL; // Все три привода и группа фактически отключены
	xDrivesReady        : BOOL; // Все приводы готовы к движению
	xDriveError         : BOOL; // Активна ошибка оси или группы осей
	xMotionBusy         : BOOL; // Одна из осей выполняет движение
	xMotionResetBusy : BOOL; // Последовательность сброса группы и осей ещё выполняется
	tSoftMotionResetTimeout : TIME := T#30S; // Предел одной принятой попытки сброса
	xSingleAxisMotionBusy : BOOL; // Один из FB_AXIS владеет осью; групповое движение запускать нельзя
	xPointCheckActive : BOOL; // Текущая команда принадлежит проверке сохранённой точки
	xTestAbort : BOOL; // Немедленная отмена активной команды виртуального теста
	rPointCheckSpeedPercent : REAL; // Фактическая скорость проверки 0.1..100 %
	lrGroupAccelerationFactor : LREAL := 1.0; // Общий разгон/торможение групповой траектории, 0.01..1.0
	lrGroupJerkFactor : LREAL := 1.0; // Общий jerk групповой траектории, 0.01..1.0
	tModbusStartTimeout : TIME := T#30S; // Ожидание создания транзакции внешним адаптером
	FaultRequest        : ST_ROBOT_FAULT_REQUEST; // Единый контракт диагностической инъекции
	tGripper1OpenTime   : TIME := T#500MS; // Время открытия первого захвата в модели
	tGripper1CloseTime  : TIME := T#500MS; // Время закрытия первого захвата в модели
	tGripper2OpenTime   : TIME := T#500MS; // Время открытия второго захвата в модели
	tGripper2CloseTime  : TIME := T#500MS; // Время закрытия второго захвата в модели
	tGripperChangeTime  : TIME := T#700MS; // Время смены рабочего захвата в модели

    stPoint : ARRAY [0..GVL_POINT.iPointNumber] OF ST_POINT; // Глобальная таблица точек робота

    xSimBlankAvailable : BOOL; // Начальное наличие заготовки в модели захвата

END_VAR
VAR_OUTPUT
	GripperCommand : ST_GRIPPER_COMMAND; // Команда для страницы физических выходов
	Command       : ST_ROBOT_COMMAND; // Выбранная команда текущего цикла
	ModbusCommand : ST_ROBOT_COMMAND; // Команда внешнему роботу по Modbus
	Status        : ST_ROBOT_STATUS; // Рабочие статусы робота
	Diag          : ST_ROBOT_DIAG; // Состояние автомата и активная команда
	Error         : ST_ROBOT_ERRORS; // Активные и последние ошибки
	GripperDiag   : ST_GRIPPER_DIAG; // Диагностика внутреннего блока захвата
	GripperError  : ST_GRIPPER_ERRORS; // Активные и последние ошибки захвата
	FaultStatus : ST_ROBOT_FAULT_STATUS; // Сводное состояние инжекторов робота
END_VAR
VAR
	fbMotionManager  : FB_MOTION_MANAGER; // Менеджер перемещения по точкам
    fbGripper        : FB_GRIPPER_SIMULATION; // Модель двухпозиционного захвата
	stGripperCommand : ST_GRIPPER_COMMAND; // Команда внутренней модели захвата

    eState        : E_ROBOT_STATE := E_ROBOT_STATE.IDLE; // Текущее состояние автомата робота
    eActiveAction : E_ROBOT_ACTION := E_ROBOT_ACTION.NONE; // Защёлкнутое действие
    eActivePoint  : E_POINT_NAME; // Защёлкнутая целевая точка
	iActiveSlot   : SINT; // Защёлкнутый слот для всей Modbus-транзакции
	uiActiveMagazineId : UINT; // Защёлкнутый магазин для всей Modbus-транзакции
	uiRobotMagazineContext : UINT; // Физический контекст магазина сохраняется между командами
	xEquipmentStopLatched : BOOL; // Робот остановлен именно аварией обслуживаемого оборудования

	xMotionExecute  : BOOL; // Запрос выполнения перемещения
	xGripperExecute : BOOL; // Запрос выполнения действия захвата
	xManualGripperRequest : BOOL; // Ручной захват разрешён независимо от состояния автомата робота
	xManualGripperOverrideExecute : BOOL; // Прямой импульс FB_GRIPPER из ERROR робота
	eManualGripperAction : E_ROBOT_ACTION; // Действие прямого ручного импульса
	xActiveManualGripper : BOOL; // Текущее действие захвата запущено вручную
	xMagazineCommandActive : BOOL; // Активная команда получена от FB_MAGAZINE
	xMagazineTargetInhibit : BOOL; // Команда входит в магазин, который меняет палеты
	rtReset               : R_TRIG; // Фронт команды сброса робота
	rtHmiDrivesEnable     : R_TRIG; // Фронт запроса включения приводов с HMI
	rtHmiDrivesDisable    : R_TRIG; // Фронт запроса отключения приводов с HMI
	rtHmiStop             : R_TRIG; // Фронт запроса остановки с HMI
	xPowerAllowed         : BOOL; // Визуальная доступность кнопки питания приводов
	xStopAllowed          : BOOL; // Визуальная доступность кнопки остановки
	xResetAllowed         : BOOL; // Визуальная доступность кнопки сброса
	xResetAccepted        : BOOL; // Общий сброс принят владельцем робота
	xExternalResetPending : BOOL; // Удерживает асинхронный Reset до подтверждения SC-500
	xExternalResetIssued  : BOOL; // Reset хотя бы один цикл был передан Modbus-адаптеру
	xSoftMotionResetPending : BOOL; // Один Reset ждёт группу, Motion и захват
	tonSoftMotionReset : TON; // Принятая попытка не может оставаться вечной
	xModbusCommandStarted : BOOL; // Текущая команда получила собственную активную транзакцию
	tonModbusStartTimeout : TON; // Защита от вечного ожидания приёма команды адаптером
	fbRobotFaultInjector  : FB_ROBOT_FAULT_INJECTOR; // Безопасная недопустимая команда робота
	xRobotFaultAllowed    : BOOL; // Владелец готов проверить тестовую команду
	uiTestBlankPayloadType : UINT;
	uiTestDetailPayloadType : UINT;
	xTestBlankPayloadPending : BOOL;
	xTestDetailPayloadPending : BOOL;

END_VAR

VAR_IN_OUT
    stMotionManager : ST_MOTION_MANAGER; // Данные менеджера движения
    GroupData       : ST_AXIS_GROUP; // Данные группы осей XYZ
    stPointManager  : ST_POINT_MANAGER; // Данные проверки точки
END_VAR

VAR CONSTANT
	ERR_ROBOT_WRONG_ACTION : DWORD := DWORD#16#0000_0001; // Недопустимое действие робота
    ERR_ROBOT_MOTION       : DWORD := DWORD#16#0000_0002; // Ошибка менеджера движения
    ERR_ROBOT_GRIPPER      : DWORD := DWORD#16#0000_0004; // Ошибка захвата
	ERR_ROBOT_MODBUS_COMM  : DWORD := DWORD#16#0000_0008; // Ошибка связи Modbus TCP
	ERR_ROBOT_STOP         : DWORD := DWORD#16#0000_0010; // Остановка команды робота
	ERR_EXTERNAL_ROBOT     : DWORD := DWORD#16#0000_0020; // Контроллер робота сообщил аварию
	WRN_RESET_EXECUTE_ACTIVE : UINT := 1; // Команда робота ещё активна
	WRN_RESET_STOP_ACTIVE    : UINT := 2; // Команда остановки ещё активна
	WRN_RESET_GLOBAL_ERROR   : UINT := 3; // Глобальная ошибка ещё активна
	WRN_RESET_MOTION_ERROR   : UINT := 4; // Ошибка менеджера движения ещё активна
	WRN_RESET_GRIPPER_ERROR  : UINT := 5; // Ошибка захвата ещё активна
	WRN_RESET_MODBUS_ERROR   : UINT := 6; // Ошибка внешнего робота ещё активна
	WRN_HMI_MANUAL_REQUIRED  : UINT := 7; // Ручная команда запрещена режимом ячейки
	WRN_DRIVES_ENABLE_ERROR  : UINT := 8; // Команда приводов отклонена владельцем Motion-слоя
	WRN_STOP_DRIVES_NOT_READY: UINT := 9; // Остановка недоступна при неготовых приводах
	WRN_SIM_ERROR_NOT_ALLOWED: UINT := 11; // Тестовая команда запрещена текущим состоянием
END_VAR

rtHmiDrivesEnable(CLK := xHmiDrivesEnable);
rtHmiDrivesDisable(CLK := xHmiDrivesDisable);
rtHmiStop(CLK := xHmiStop);

xPowerAllowed := ((NOT xDrivesOff) AND xHmiDrivesDisableAllowed)
	OR (xDrivesOff AND xHmiDrivesEnableAllowed);
xStopAllowed := xHmiStopAllowed;

IF (rtHmiDrivesEnable.Q AND NOT xHmiDrivesEnableAccepted)
OR (rtHmiDrivesDisable.Q AND NOT xHmiDrivesDisableAccepted) THEN
	IF NOT xHmiPermit THEN
		Diag.stWarning.uiCode := WRN_HMI_MANUAL_REQUIRED;
	ELSE
		Diag.stWarning.uiCode := WRN_DRIVES_ENABLE_ERROR;
	END_IF;
	Diag.stWarning.udiSequence := Diag.stWarning.udiSequence + UDINT#1;
	IF Diag.stWarning.udiSequence = UDINT#0 THEN
		Diag.stWarning.udiSequence := UDINT#1;
	END_IF;
END_IF;

IF rtHmiStop.Q
AND NOT xHmiStopAccepted THEN
	IF NOT xHmiPermit THEN
		Diag.stWarning.uiCode := WRN_HMI_MANUAL_REQUIRED;
	ELSE
		Diag.stWarning.uiCode := WRN_STOP_DRIVES_NOT_READY;
	END_IF;
	Diag.stWarning.udiSequence := Diag.stWarning.udiSequence + UDINT#1;
	IF Diag.stWarning.udiSequence = UDINT#0 THEN
		Diag.stWarning.udiSequence := UDINT#1;
	END_IF;
END_IF;

// Команды по умолчанию
xMotionExecute := FALSE;
xGripperExecute := FALSE;
xManualGripperRequest := FALSE;
xManualGripperOverrideExecute := FALSE;
xMagazineCommandActive := FALSE;
xMagazineTargetInhibit := FALSE;

Command.xExecute := FALSE;
Command.xStop := FALSE;
Command.xReset := FALSE;
Command.eAction := E_ROBOT_ACTION.NONE;
Command.eSetPoint := E_POINT_NAME.NONE;
Command.iActiveSlot := 0;
Command.uiMagazineId := UINT#0;

ModbusCommand.xExecute := FALSE;
ModbusCommand.xStop := FALSE;
ModbusCommand.xReset := FALSE;
ModbusCommand.eAction := E_ROBOT_ACTION.NONE;
ModbusCommand.eSetPoint := E_POINT_NAME.NONE;
ModbusCommand.iActiveSlot := 0;
ModbusCommand.uiMagazineId := UINT#0;

//Определяем какой режим работы активен
IF NOT xManual THEN
	IF stCellCommand.xExecute OR stCellCommand.xStop THEN
		Command := stCellCommand;
	ELSIF stMachine_1_Command.xExecute OR stMachine_1_Command.xStop THEN
		Command := stMachine_1_Command;
	ELSIF stMachine_2_Command.xExecute OR stMachine_2_Command.xStop THEN
		Command := stMachine_2_Command;
	ELSIF stMachine_3_Command.xExecute OR stMachine_3_Command.xStop THEN
		Command := stMachine_3_Command;
	ELSIF stMagazineCommand.xExecute OR stMagazineCommand.xStop THEN
		Command := stMagazineCommand;
		xMagazineCommandActive := TRUE;
	END_IF;
ELSE
	IF stMagazineCommand.xExecute OR stMagazineCommand.xStop THEN
		Command := stMagazineCommand;
		xMagazineCommandActive := TRUE;
	ELSE
		Command := stHmiCommand;
	END_IF;
END_IF;

// Смена палет блокирует автоматические команды и операции FB_MAGAZINE
// с этим магазином. Ручная точка HMI не зависит от состояния магазина.
IF (NOT xManual OR xMagazineCommandActive)
AND (Command.uiMagazineId >= UINT#1) AND (Command.uiMagazineId <= UINT#2) THEN
	IF axMagazineExchangeInProgress[Command.uiMagazineId] THEN
		IF (Command.eSetPoint = E_POINT_NAME.MAGAZINE_SAFE)
		OR (Command.eSetPoint = E_POINT_NAME.MAGAZINE_CHANGE)
		OR (Command.eSetPoint = E_POINT_NAME.MAGAZINE_IN_SLOT) THEN
			xMagazineTargetInhibit := TRUE;
		END_IF;
	END_IF;
END_IF;

// Abort теста имеет приоритет над любым владельцем, включая ручную подготовку
// сценария, когда команда ячейки обычно не участвует в выборе.
IF xTestAbort THEN
	Command.xExecute := FALSE;
	Command.xStop := TRUE;
END_IF;

// Уже принятую внешним контроллером команду не прерываем. Запрет действует
// только в IDLE, то есть перед началом следующего высокоуровневого действия.
IF xMode
AND xExternalCommandInhibit
AND (eState = E_ROBOT_STATE.IDLE) THEN
	Command.xExecute := FALSE;
END_IF;

IF xMagazineTargetInhibit AND (eState = E_ROBOT_STATE.IDLE) THEN
	Command.xExecute := FALSE;
END_IF;

// Внешний Stop — самостоятельная приоритетная команда. Он должен дойти до
// адаптера и тогда, когда FB_ROBOT уже защёлкнул ERROR после общей остановки.
IF xMode
AND (xHmiStopAccepted
	OR Command.xStop
	OR (xGlobalError AND stModbusStatus.xBusy)) THEN
	ModbusCommand.xStop := TRUE;
END_IF;

// Класс ошибки определяет оборудование-владелец. FB_ROBOT только выполняет
// зависимую реакцию: активное действие останавливает, неподвижный робот сразу
// переводит в ERROR без бессмысленной команды Stop.
IF xEquipmentStopRequired
AND (eState <> E_ROBOT_STATE.ERROR) THEN
	xEquipmentStopLatched := TRUE;
	IF (eState = E_ROBOT_STATE.MOTION)
	OR (eState = E_ROBOT_STATE.GRIPPER)
	OR (eState = E_ROBOT_STATE.MODBUS) THEN
		Command.xStop := TRUE;
	ELSE
		Error.dwErrorActive := Error.dwErrorActive OR ERR_ROBOT_STOP;
		eState := E_ROBOT_STATE.ERROR;
	END_IF;
END_IF;

// RunRobot уже выполнил все PLC-проверки и передал Execute только принятой
// ручной команде. Захват остаётся независимым от состояния осей и робота.
IF xManual AND stHmiCommand.xExecute THEN
	CASE stHmiCommand.eAction OF
		E_ROBOT_ACTION.UNCLAMP_1,
		E_ROBOT_ACTION.CLAMP_1,
		E_ROBOT_ACTION.UNCLAMP_2,
		E_ROBOT_ACTION.CLAMP_2,
		E_ROBOT_ACTION.ROTATE_TO_BLANK,
		E_ROBOT_ACTION.ROTATE_TO_DETAIL:
			xManualGripperRequest := TRUE;
	END_CASE;
END_IF;

// Готовность сброса рассчитывается после выбора актуального владельца команды.
// Ошибки вложенных FB считаются сбрасываемыми только после снятия удерживаемого
// источника и публикации их собственного xResetAllowed.
rtReset(CLK := xReset);
xResetAllowed := xHmiPermit
	AND NOT xSoftMotionResetPending
	AND NOT xExternalResetPending
	AND (NOT xMode OR NOT stModbusStatus.xResetBusy)
	AND (NOT xGlobalError OR xManualRecoveryAllowed)
	AND NOT Command.xExecute
	AND NOT Command.xStop
	AND NOT xMotionBusy
	AND (NOT xMode OR stModbusStatus.xCommunicationAlive)
	AND (xDriveError
		OR (eState = E_ROBOT_STATE.ERROR)
		OR (NOT xMode AND stMotionManager.Status.xError)
		OR (NOT xMode AND fbGripper.Status.xError)
		OR (xMode AND xModbusError))
	AND (xMode OR NOT stMotionManager.Status.xError
		OR FaultStatus.stPoint.xResetAllowed)
	AND (xMode OR NOT fbGripper.Status.xError
		OR FaultStatus.stGripper.xResetAllowed);
xResetAccepted := rtReset.Q AND xResetAllowed;
// Общий Reset запускает Motion-сброс раньше FB_ROBOT. Если группа была в
// ErrorStop, одноцикловый импульс уже закончится к моменту её восстановления;
// защёлкиваем намерение оператора до исчезновения первичной Motion-ошибки.
IF xMode THEN
	xSoftMotionResetPending := FALSE;
ELSIF xResetAccepted
AND (eState = E_ROBOT_STATE.ERROR) THEN
	xSoftMotionResetPending := TRUE;
END_IF;
IF xMode AND xResetAccepted THEN
	xExternalResetPending := TRUE;
	xExternalResetIssued := FALSE;
ELSIF NOT xMode THEN
	xExternalResetPending := FALSE;
	xExternalResetIssued := FALSE;
END_IF;

tonSoftMotionReset(IN := xSoftMotionResetPending, PT := tSoftMotionResetTimeout);
IF xSoftMotionResetPending AND NOT xResetAccepted
AND (tonSoftMotionReset.Q
	OR xTestAbort OR NOT xHmiPermit OR Command.xExecute OR Command.xStop
	OR (xGlobalError AND NOT xManualRecoveryAllowed)
	OR (xDriveError AND NOT xMotionResetBusy)
	OR (fbGripper.Status.xError AND NOT FaultStatus.stGripper.xResetAllowed)
	OR (stMotionManager.Status.xError AND NOT FaultStatus.stPoint.xResetAllowed)) THEN
	xSoftMotionResetPending := FALSE;
	IF fbGripper.Status.xError THEN
		Diag.stWarning.uiCode := WRN_RESET_GRIPPER_ERROR;
	ELSE
		Diag.stWarning.uiCode := WRN_RESET_MOTION_ERROR;
	END_IF;
	Diag.stWarning.udiSequence := Diag.stWarning.udiSequence + UDINT#1;
	IF Diag.stWarning.udiSequence = UDINT#0 THEN Diag.stWarning.udiSequence := UDINT#1; END_IF;
END_IF;

// После неуспешной попытки адаптер публикует явный результат. Снимаем уровень,
// чтобы следующее осознанное нажатие Reset снова дошло до его R_TRIG.
IF xExternalResetPending AND xExternalResetIssued AND NOT xResetAccepted
AND (stModbusStatus.xResetFailed OR NOT stModbusStatus.xCommunicationAlive
	OR xTestAbort OR Command.xStop OR NOT xHmiPermit
	OR (xGlobalError AND NOT xManualRecoveryAllowed)) THEN
	xExternalResetPending := FALSE;
	xExternalResetIssued := FALSE;
	Diag.stWarning.uiCode := WRN_RESET_MODBUS_ERROR;
	Diag.stWarning.udiSequence := Diag.stWarning.udiSequence + UDINT#1;
	IF Diag.stWarning.udiSequence = UDINT#0 THEN Diag.stWarning.udiSequence := UDINT#1; END_IF;
END_IF;

// Недопустимое действие проверяется в IDLE до запуска Motion или захвата.
xRobotFaultAllowed := (eState = E_ROBOT_STATE.IDLE)
	AND NOT Command.xExecute
	AND NOT Command.xStop
	AND NOT xMode
	AND NOT xGlobalError
	AND NOT xDriveError
	AND (Error.dwErrorActive = DWORD#0)
	AND NOT stMotionManager.Status.xError
	AND NOT fbGripper.Status.xError;

fbRobotFaultInjector(
	Request := FaultRequest,
	xOwnerAllowed := xRobotFaultAllowed
);
FaultStatus.stRobot := fbRobotFaultInjector.Status;

IF fbRobotFaultInjector.Status.xRejected THEN
	Diag.stWarning.uiCode := WRN_SIM_ERROR_NOT_ALLOWED;
	Diag.stWarning.udiSequence := Diag.stWarning.udiSequence + UDINT#1;
	IF Diag.stWarning.udiSequence = UDINT#0 THEN
		Diag.stWarning.udiSequence := UDINT#1;
	END_IF;
END_IF;

IF fbRobotFaultInjector.xWrongAction THEN
	Command.xExecute := TRUE;
	Command.xStop := FALSE;
	Command.eAction := E_ROBOT_ACTION.NONE;
	Command.eSetPoint := E_POINT_NAME.NONE;
END_IF;

Command.xReset := xResetAccepted;

IF rtReset.Q
AND ((eState = E_ROBOT_STATE.ERROR) OR xDriveError)
AND NOT xResetAccepted THEN
	IF NOT xHmiPermit THEN
		Diag.stWarning.uiCode := WRN_HMI_MANUAL_REQUIRED;
	ELSIF eState <> E_ROBOT_STATE.ERROR THEN
		// Ошибку Motion-слоя сбрасывают оси и группа тем же общим импульсом.
		Diag.stWarning.uiCode := UINT#0;
    ELSIF Command.xExecute THEN
        Diag.stWarning.uiCode := WRN_RESET_EXECUTE_ACTIVE;
    ELSIF Command.xStop THEN
        Diag.stWarning.uiCode := WRN_RESET_STOP_ACTIVE;
    ELSIF xGlobalError AND NOT xManualRecoveryAllowed THEN
        Diag.stWarning.uiCode := WRN_RESET_GLOBAL_ERROR;
    ELSIF stMotionManager.Status.xError
	OR (NOT xMode AND xDriveError) THEN
        Diag.stWarning.uiCode := WRN_RESET_MOTION_ERROR;
    ELSIF fbGripper.Status.xError THEN
        Diag.stWarning.uiCode := WRN_RESET_GRIPPER_ERROR;
    ELSIF xModbusError THEN
        Diag.stWarning.uiCode := WRN_RESET_MODBUS_ERROR;
    ELSE
        Diag.stWarning.uiCode := UINT#0;
    END_IF;

    IF Diag.stWarning.uiCode <> UINT#0 THEN
        Diag.stWarning.udiSequence := Diag.stWarning.udiSequence + UDINT#1;
        IF Diag.stWarning.udiSequence = UDINT#0 THEN
            Diag.stWarning.udiSequence := UDINT#1;
        END_IF;
    END_IF;
END_IF;

// =====================================================
// Автомат FB_ROBOT
// =====================================================

// Таймаут исполнения принадлежит FB_ROBOT_MODBUS, но до создания активной
// транзакции его TON ещё не работает. Отдельно ограничиваем фазу ожидания Busy.
tonModbusStartTimeout(
	IN := xMode
		AND (eState = E_ROBOT_STATE.MODBUS)
		AND NOT xModbusCommandStarted,
	PT := tModbusStartTimeout
);

// Ошибка оси или группы является первопричиной в Motion-слое и отдельной
// каскадной ошибкой робота для его публичного статуса и журнала.
IF NOT xMode AND xDriveError THEN
	Error.dwErrorActive := Error.dwErrorActive OR ERR_ROBOT_MOTION;
	eState := E_ROBOT_STATE.ERROR;
ELSIF NOT xMode AND stMotionManager.Status.xError THEN
	// Отмена задания при ручном I/O не скрывает аварию вложенного владельца.
	Error.dwErrorActive := Error.dwErrorActive OR ERR_ROBOT_MOTION;
	eState := E_ROBOT_STATE.ERROR;
ELSIF NOT xMode AND fbGripper.Status.xError THEN
	Error.dwErrorActive := Error.dwErrorActive OR ERR_ROBOT_GRIPPER;
	eState := E_ROBOT_STATE.ERROR;
ELSIF xMode AND xModbusError THEN
	IF stModbusStatus.xRobotAlarm THEN
		Error.dwErrorActive := Error.dwErrorActive OR ERR_EXTERNAL_ROBOT;
	ELSE
		Error.dwErrorActive := Error.dwErrorActive OR ERR_ROBOT_MODBUS_COMM;
	END_IF;
	eState := E_ROBOT_STATE.ERROR;
END_IF;

CASE eState OF

    E_ROBOT_STATE.IDLE:

        Status.xBusy := FALSE;
        Status.xDone := FALSE;
        Status.xError := FALSE;

        IF Command.xExecute THEN
            eActiveAction := Command.eAction;
            eActivePoint := Command.eSetPoint;
			iActiveSlot := Command.iActiveSlot;
			uiActiveMagazineId := Command.uiMagazineId;
			IF (Command.uiMagazineId >= UINT#1)
			AND (Command.uiMagazineId <= UINT#2)
			AND (Command.eAction = E_ROBOT_ACTION.MOVE_TO_POINT)
			AND ((Command.eSetPoint = E_POINT_NAME.MAGAZINE_IN_SLOT)
				OR (Command.eSetPoint = E_POINT_NAME.MAGAZINE_CHANGE)) THEN
				uiRobotMagazineContext := Command.uiMagazineId;
			END_IF;

            IF xMode THEN
				xModbusCommandStarted := FALSE;
				eState := E_ROBOT_STATE.MODBUS;

            ELSE
                CASE Command.eAction OF

                    E_ROBOT_ACTION.MOVE_TO_POINT:
                        // CODESYS переводит группу в ошибку, если GroupMoving
                        // запускается при активном single-axis FB. Команда
                        // остаётся в IDLE до освобождения всех FB_AXIS.
                        IF xDrivesReady AND NOT xMotionBusy THEN
                            eState := E_ROBOT_STATE.MOTION;
                        END_IF;

                    E_ROBOT_ACTION.UNCLAMP_1,
                    E_ROBOT_ACTION.CLAMP_1,
                    E_ROBOT_ACTION.UNCLAMP_2,
                    E_ROBOT_ACTION.CLAMP_2,
                    E_ROBOT_ACTION.ROTATE_TO_BLANK,
                    E_ROBOT_ACTION.ROTATE_TO_DETAIL:
						xActiveManualGripper := xManualGripperRequest;
                        eState := E_ROBOT_STATE.GRIPPER;

                ELSE
                    Error.dwErrorActive :=
                        Error.dwErrorActive OR ERR_ROBOT_WRONG_ACTION;

                    eState := E_ROBOT_STATE.ERROR;
                END_CASE;
            END_IF;
        END_IF;


    E_ROBOT_STATE.MOTION:

        Status.xBusy := TRUE;
        xMotionExecute := NOT xSingleAxisMotionBusy;

		IF xHmiStopAccepted OR Command.xStop THEN
			// Операторский Stop отменяет действие штатно. Stop от оборудования
			// дополнительно защёлкивает зависимую ошибку робота.
            xMotionExecute := FALSE;
            Status.xBusy := FALSE;
            Status.xDone := FALSE;
            eActiveAction := E_ROBOT_ACTION.NONE;
            eActivePoint := E_POINT_NAME.NONE;
			IF xEquipmentStopRequired THEN
				Error.dwErrorActive := Error.dwErrorActive OR ERR_ROBOT_STOP;
				eState := E_ROBOT_STATE.ERROR;
			ELSE
				eState := E_ROBOT_STATE.IDLE;
			END_IF;

        ELSIF xGlobalError THEN
            Error.dwErrorActive := Error.dwErrorActive OR ERR_ROBOT_STOP;
            eState := E_ROBOT_STATE.ERROR;

        ELSIF stMotionManager.Status.xError THEN
            Error.dwErrorActive := Error.dwErrorActive OR ERR_ROBOT_MOTION;
            eState := E_ROBOT_STATE.ERROR;

		ELSIF stMotionManager.Status.xDone THEN
			IF (eActiveAction = E_ROBOT_ACTION.MOVE_TO_POINT)
			AND (eActivePoint <> E_POINT_NAME.MAGAZINE_IN_SLOT)
			AND (eActivePoint <> E_POINT_NAME.MAGAZINE_CHANGE) THEN
				uiRobotMagazineContext := UINT#0;
			END_IF;
            eState := E_ROBOT_STATE.DONE;
        END_IF;


	E_ROBOT_STATE.GRIPPER:

        Status.xBusy := TRUE;
        xGripperExecute := TRUE;

		IF xTestAbort THEN
			xGripperExecute := FALSE;
			Status.xBusy := FALSE;
			Status.xDone := FALSE;
			xActiveManualGripper := FALSE;
			eActiveAction := E_ROBOT_ACTION.NONE;
			eActivePoint := E_POINT_NAME.NONE;
			eState := E_ROBOT_STATE.IDLE;

		ELSIF xEquipmentStopRequired THEN
			xGripperExecute := FALSE;
			Error.dwErrorActive := Error.dwErrorActive OR ERR_ROBOT_STOP;
			eState := E_ROBOT_STATE.ERROR;

		ELSIF xGlobalError AND NOT xActiveManualGripper THEN
            Error.dwErrorActive := Error.dwErrorActive OR ERR_ROBOT_STOP;
            eState := E_ROBOT_STATE.ERROR;

        ELSIF fbGripper.Status.xError THEN
            Error.dwErrorActive := Error.dwErrorActive OR ERR_ROBOT_GRIPPER;
            eState := E_ROBOT_STATE.ERROR;

        ELSIF fbGripper.Status.xDone THEN
			xActiveManualGripper := FALSE;
            eState := E_ROBOT_STATE.DONE;
        END_IF;


	E_ROBOT_STATE.DONE:

        Status.xBusy := FALSE;
        Status.xDone := TRUE;

        IF NOT xMode THEN
        CASE eActiveAction OF

            E_ROBOT_ACTION.MOVE_TO_POINT:
                xMotionExecute := TRUE;

            E_ROBOT_ACTION.UNCLAMP_1,
            E_ROBOT_ACTION.CLAMP_1,
            E_ROBOT_ACTION.UNCLAMP_2,
            E_ROBOT_ACTION.CLAMP_2,
            E_ROBOT_ACTION.ROTATE_TO_BLANK,
            E_ROBOT_ACTION.ROTATE_TO_DETAIL:
                xGripperExecute := TRUE;

        END_CASE;
        END_IF;

		IF NOT Command.xExecute THEN
			// Владелец уже снял Execute: в этом же цикле погасить запрос
			// вложенному FB до очистки action/point. Иначе при быстром
			// SoftMotion движении один скан уходил как Execute=TRUE + point=NONE,
			// а FB_MOTION_MANAGER закономерно валил нулевую точку.
			xMotionExecute := FALSE;
			xGripperExecute := FALSE;
            Status.xDone := FALSE;
			xModbusCommandStarted := FALSE;
            eActiveAction := E_ROBOT_ACTION.NONE;
			eActivePoint := E_POINT_NAME.NONE;
			iActiveSlot := SINT#0;
			uiActiveMagazineId := UINT#0;
			eState := E_ROBOT_STATE.IDLE;
        END_IF;


	E_ROBOT_STATE.MODBUS:
		Status.xBusy := TRUE;
		// Execute — импульс от владельца команды. Адаптер Modbus может
		// быть занят FC03/FC16 дольше этого импульса. Поэтому до терминального
		// ответа передаём защёлкнутые action/point/slot, а не уже снятый Command.
		ModbusCommand.xExecute := TRUE;
		ModbusCommand.eAction := eActiveAction;
		ModbusCommand.eSetPoint := eActivePoint;
		ModbusCommand.iActiveSlot := iActiveSlot;
		ModbusCommand.uiMagazineId := uiActiveMagazineId;
		IF xModbusBusy THEN
			xModbusCommandStarted := TRUE;
		END_IF;

		IF xTestAbort THEN
			ModbusCommand.xStop := TRUE;
			IF NOT stModbusStatus.xBusy THEN
				Status.xBusy := FALSE;
				Status.xDone := FALSE;
				xModbusCommandStarted := FALSE;
				eActiveAction := E_ROBOT_ACTION.NONE;
				eActivePoint := E_POINT_NAME.NONE;
				iActiveSlot := SINT#0;
				uiActiveMagazineId := UINT#0;
				eState := E_ROBOT_STATE.IDLE;
			END_IF;
		ELSIF Command.xStop OR xHmiStopAccepted OR xGlobalError THEN
			ModbusCommand.xStop := TRUE;
			Error.dwErrorActive := Error.dwErrorActive OR ERR_ROBOT_STOP;
			eState := E_ROBOT_STATE.ERROR;
		ELSIF xModbusError THEN
			IF stModbusStatus.xRobotAlarm THEN
				Error.dwErrorActive := Error.dwErrorActive OR ERR_EXTERNAL_ROBOT;
			ELSE
				Error.dwErrorActive := Error.dwErrorActive OR ERR_ROBOT_MODBUS_COMM;
			END_IF;
			eState := E_ROBOT_STATE.ERROR;
		ELSIF tonModbusStartTimeout.Q THEN
			// Адаптер не создал собственную транзакцию: не оставляем публичный
			// xBusy висеть бесконечно без CommandSeq и физического движения.
			ModbusCommand.xExecute := FALSE;
			Error.dwErrorActive := Error.dwErrorActive OR ERR_ROBOT_MODBUS_COMM;
			eState := E_ROBOT_STATE.ERROR;
		ELSIF xModbusCommandStarted AND xModbusDone THEN
			IF (eActiveAction = E_ROBOT_ACTION.MOVE_TO_POINT)
			AND (eActivePoint <> E_POINT_NAME.MAGAZINE_IN_SLOT)
			AND (eActivePoint <> E_POINT_NAME.MAGAZINE_CHANGE) THEN
				uiRobotMagazineContext := UINT#0;
			END_IF;
			eState := E_ROBOT_STATE.DONE;
		END_IF;


    E_ROBOT_STATE.ERROR:

        Status.xBusy := FALSE;
        Status.xDone := FALSE;
        Status.xError := TRUE;

		// Ошибка координатного робота не блокирует независимый ручной захват.
		// Собственная ошибка FB_GRIPPER по-прежнему требует штатного сброса.
		IF NOT xMode AND xManualGripperRequest AND NOT fbGripper.Status.xError THEN
			xManualGripperOverrideExecute := TRUE;
			eManualGripperAction := stHmiCommand.eAction;
		END_IF;

		// В Modbus-режиме входной Reset только защёлкивает запрос для адаптера.
		// Локальную ошибку можно снять лишь после подтверждённого исчезновения
		// внешней аварии; иначе xExternalResetPending очистится до записи 1004.
		IF ((NOT xMode AND (xResetAccepted OR xSoftMotionResetPending))
			OR (xMode
				AND xExternalResetPending
				AND xExternalResetIssued
				AND stModbusStatus.xResetDone
				AND NOT xModbusError
				AND NOT stModbusStatus.xBusy
				AND (stModbusStatus.uiExecutionState =
					TO_UINT(E_ROBOT_MODBUS_EXECUTION_STATE.IDLE))))
        AND NOT Command.xExecute
        AND NOT Command.xStop
        AND (NOT xGlobalError OR xManualRecoveryAllowed)
		AND (xMode OR NOT stMotionManager.Status.xError)
		AND (xMode OR NOT xDriveError)
		AND (xMode OR NOT fbGripper.Status.xError)
		AND (NOT xMode OR stModbusStatus.xCommunicationAlive) THEN

			Error.dwErrorLast := Error.dwErrorActive;
			Error.dwErrorActive := DWORD#0;
            Status.xError := FALSE;
			xExternalResetPending := FALSE;
			xExternalResetIssued := FALSE;
			xSoftMotionResetPending := FALSE;
			xModbusCommandStarted := FALSE;
			xActiveManualGripper := FALSE;
			xEquipmentStopLatched := FALSE;
            eActiveAction := E_ROBOT_ACTION.NONE;
			eActivePoint := E_POINT_NAME.NONE;
			iActiveSlot := SINT#0;
			uiActiveMagazineId := UINT#0;
			eState := E_ROBOT_STATE.IDLE;
        END_IF;

END_CASE;

IF xMode AND xExternalResetPending THEN
	ModbusCommand.xReset := TRUE;
	xExternalResetIssued := TRUE;
END_IF;

// =====================================================
// Формирование команды FB_MOTION_MANAGER
// =====================================================

stMotionManager.Command.xExecute := NOT xMode AND xMotionExecute;
stMotionManager.Command.eTargetPoint := eActivePoint;
stMotionManager.Command.xReset := NOT xMode AND xResetAccepted;
stMotionManager.Command.xStop := NOT xMode AND (xHmiStopAccepted OR Command.xStop);
stMotionManager.Command.xGlobalError :=
    (NOT xMode AND xGlobalError AND NOT xManualRecoveryAllowed);


// =====================================================
// Вызов FB_MOTION_MANAGER
// =====================================================

fbMotionManager(
    stPoint := stPoint,
    xReset := NOT xMode AND xResetAccepted,
	FaultRequest := FaultRequest.stPoint,
	xSpeedFactorOverride := xPointCheckActive,
	lrSpeedFactorOverride := REAL_TO_LREAL(rPointCheckSpeedPercent) / 100.0,
	lrAccelerationFactor := lrGroupAccelerationFactor,
	lrJerkFactor := lrGroupJerkFactor,
    stMotionManager := stMotionManager,
    GroupData := GroupData,
    stPointManager := stPointManager
);
FaultStatus.stPoint := fbMotionManager.FaultStatus;


// =====================================================
// Вызов FB_GRIPPER
// =====================================================

stGripperCommand.xExecute := NOT xMode
	AND (xGripperExecute OR xManualGripperOverrideExecute);
stGripperCommand.xReset := NOT xMode AND xResetAccepted;
stGripperCommand.xGripper1Open := fbGripper.Status.xGripper1Open;
stGripperCommand.xGripper2Open := fbGripper.Status.xGripper2Open;
stGripperCommand.xRotateToDetail := fbGripper.Status.xRotatedToDetail;
IF xManualGripperOverrideExecute THEN
	stGripperCommand.eAction := eManualGripperAction;
ELSE
	stGripperCommand.eAction := eActiveAction;
END_IF;
CASE stGripperCommand.eAction OF
	E_ROBOT_ACTION.UNCLAMP_1: stGripperCommand.xGripper1Open := TRUE;
	E_ROBOT_ACTION.CLAMP_1: stGripperCommand.xGripper1Open := FALSE;
	E_ROBOT_ACTION.UNCLAMP_2: stGripperCommand.xGripper2Open := TRUE;
	E_ROBOT_ACTION.CLAMP_2: stGripperCommand.xGripper2Open := FALSE;
	E_ROBOT_ACTION.ROTATE_TO_BLANK: stGripperCommand.xRotateToDetail := FALSE;
	E_ROBOT_ACTION.ROTATE_TO_DETAIL: stGripperCommand.xRotateToDetail := TRUE;
END_CASE;

GripperCommand := stGripperCommand;
fbGripper(
	xUsePhysicalFeedback := xUsePhysicalGripperFeedback AND NOT xMode,
	xPhysicalIoReady := xPhysicalGripperIoReady,
	PhysicalFeedback := stPhysicalGripperFeedback,
	tPhysicalActionTimeout := tPhysicalGripperActionTimeout,
	// Положение и захваты робота не подменяются записью сценария: runner
	// приводит их в нужное состояние штатными командами.
	xTestInitialize := FALSE,
	auiTestContent := auiTestGripperContent,
	uiTestOrientation := uiTestOrientation,
	Command := stGripperCommand,
	FaultRequest := FaultRequest.stGripper,
	xSimulationAccelerationEnable := xSimulationAccelerationEnable,
	uiSimulationTimeFactor := uiSimulationTimeFactor,
	tGripper1OpenTime := tGripper1OpenTime,
	tGripper1CloseTime := tGripper1CloseTime,
	tGripper2OpenTime := tGripper2OpenTime,
	tGripper2CloseTime := tGripper2CloseTime,
	tRotateTime := tGripperChangeTime,
	Diag => GripperDiag,
	Error => GripperError
);
FaultStatus.stGripper := fbGripper.FaultStatus;

IF xTestInitialize THEN
	uiTestBlankPayloadType := auiTestGripperType[1];
	uiTestDetailPayloadType := auiTestGripperType[2];
	xTestBlankPayloadPending := auiTestGripperContent[1] = UINT#1;
	xTestDetailPayloadPending := auiTestGripperContent[2] = UINT#2;
	uiRobotMagazineContext := UINT#0;
	xEquipmentStopLatched := FALSE;
	xSoftMotionResetPending := FALSE;
END_IF;


// =====================================================
// Общие статусы
// =====================================================

IF xMode THEN
	CASE stModbusStatus.uiCurrentPoint OF
		10: Status.eCurrentPoint := E_POINT_NAME.MACHINE_1_ABOVE;
		11: Status.eCurrentPoint := E_POINT_NAME.MACHINE_1_INSIDE;
		12: Status.eCurrentPoint := E_POINT_NAME.MACHINE_1_CHUCK_APROACH;
		13: Status.eCurrentPoint := E_POINT_NAME.MACHINE_1_CHUCK_POSITION;
		14: Status.eCurrentPoint := E_POINT_NAME.MACHINE_2_ABOVE;
		15: Status.eCurrentPoint := E_POINT_NAME.MACHINE_2_INSIDE;
		16: Status.eCurrentPoint := E_POINT_NAME.MACHINE_2_CHUCK_APROACH;
		17: Status.eCurrentPoint := E_POINT_NAME.MACHINE_2_CHUCK_POSITION;
		18: Status.eCurrentPoint := E_POINT_NAME.MACHINE_3_ABOVE;
		19: Status.eCurrentPoint := E_POINT_NAME.MACHINE_3_INSIDE;
		20: Status.eCurrentPoint := E_POINT_NAME.MACHINE_3_CHUCK_APROACH;
		21: Status.eCurrentPoint := E_POINT_NAME.MACHINE_3_CHUCK_POSITION;
		22: Status.eCurrentPoint := E_POINT_NAME.HOME_SAFETY;
		23: Status.eCurrentPoint := E_POINT_NAME.MAGAZINE_SAFE;
		24: Status.eCurrentPoint := E_POINT_NAME.MAGAZINE_CHANGE;
		25: Status.eCurrentPoint := E_POINT_NAME.MAGAZINE_IN_SLOT;
	ELSE
		Status.eCurrentPoint := E_POINT_NAME.NONE;
	END_CASE;
	Status.xGripper1Open := (stModbusStatus.uiGripperStatus AND UINT#16#0001) <> UINT#0;
	Status.xGripper1Closed := (stModbusStatus.uiGripperStatus AND UINT#16#0002) <> UINT#0;
	Status.xGripper2Open := (stModbusStatus.uiGripperStatus AND UINT#16#0004) <> UINT#0;
	Status.xGripper2Closed := (stModbusStatus.uiGripperStatus AND UINT#16#0008) <> UINT#0;
	Status.xRotatedToBlank := (stModbusStatus.uiGripperStatus AND UINT#16#0010) <> UINT#0;
	Status.xRotatedToDetail := (stModbusStatus.uiGripperStatus AND UINT#16#0020) <> UINT#0;
ELSE
	Status.eCurrentPoint := stMotionManager.Status.eCurrentPoint;
	Status.xGripper1Open := fbGripper.Status.xGripper1Open;
	Status.xGripper1Closed := fbGripper.Status.xGripper1Closed;
	Status.xGripper2Open := fbGripper.Status.xGripper2Open;
	Status.xGripper2Closed := fbGripper.Status.xGripper2Closed;
	Status.xRotatedToBlank := fbGripper.Status.xRotatedToBlank;
	Status.xRotatedToDetail := fbGripper.Status.xRotatedToDetail;
END_IF;

Status.xBlankAvailable := Status.xGripper1Closed;
Status.xDetailAvailable := Status.xGripper2Closed;
IF Status.xGripper1Open THEN
	Status.uiBlankPayloadType := UINT#0;
	IF NOT xTestBlankPayloadPending THEN
		uiTestBlankPayloadType := UINT#0;
	END_IF;
ELSIF Status.xGripper1Closed THEN
	// Во время загрузки тестового сценария его тип относится к уже заданному
	// содержимому захвата и имеет приоритет над метаданными предыдущего цикла.
	IF xTestBlankPayloadPending
	AND (uiTestBlankPayloadType >= UINT#1)
	AND (uiTestBlankPayloadType <= UINT#3) THEN
		Status.uiBlankPayloadType := uiTestBlankPayloadType;
	ELSIF (uiBlankPayloadType >= UINT#1) AND (uiBlankPayloadType <= UINT#3) THEN
		Status.uiBlankPayloadType := uiBlankPayloadType;
		uiTestBlankPayloadType := uiBlankPayloadType;
	ELSIF (uiTestBlankPayloadType >= UINT#1)
	AND (uiTestBlankPayloadType <= UINT#3) THEN
		Status.uiBlankPayloadType := uiTestBlankPayloadType;
	ELSE
		Status.uiBlankPayloadType := UINT#0;
	END_IF;
	xTestBlankPayloadPending := FALSE;
END_IF;
IF Status.xGripper2Open THEN
	Status.uiDetailPayloadType := UINT#0;
	IF NOT xTestDetailPayloadPending THEN
		uiTestDetailPayloadType := UINT#0;
	END_IF;
ELSIF Status.xGripper2Closed THEN
	IF xTestDetailPayloadPending
	AND (uiTestDetailPayloadType >= UINT#1)
	AND (uiTestDetailPayloadType <= UINT#3) THEN
		Status.uiDetailPayloadType := uiTestDetailPayloadType;
	ELSIF (uiDetailPayloadType >= UINT#1) AND (uiDetailPayloadType <= UINT#3) THEN
		Status.uiDetailPayloadType := uiDetailPayloadType;
		uiTestDetailPayloadType := uiDetailPayloadType;
	ELSIF (uiTestDetailPayloadType >= UINT#1)
	AND (uiTestDetailPayloadType <= UINT#3) THEN
		Status.uiDetailPayloadType := uiTestDetailPayloadType;
	ELSE
		Status.uiDetailPayloadType := UINT#0;
	END_IF;
	xTestDetailPayloadPending := FALSE;
END_IF;
Status.xPowerAllowed := xPowerAllowed;
Status.xStopAllowed := xStopAllowed;
Status.xResetAllowed := xResetAllowed;
Status.uiMagazineContext := uiRobotMagazineContext;

Diag.eState := eState;
Diag.eActiveAction := eActiveAction;
Diag.eActivePoint := eActivePoint;
Error.dwAlarmActive := Error.dwErrorActive;
Status.xExternalError := ((Error.dwErrorActive AND (ERR_ROBOT_MOTION OR ERR_ROBOT_GRIPPER)) <> DWORD#0)
	OR xEquipmentStopLatched;

IF Error.dwErrorActive <> DWORD#0 THEN
	Error.dwErrorLast := Error.dwErrorActive;
END_IF;

Error.stErrorActive := UpdateErrorView(dwError := Error.dwErrorActive);
Error.stErrorLast := UpdateErrorView(dwError := Error.dwErrorLast);
FaultStatus.stRobot.xResetAllowed := Status.xResetAllowed
	AND NOT FaultStatus.stRobot.xBusy;

METHOD UpdateErrorView : ST_ROBOT_ERROR
VAR_INPUT
	dwError : DWORD; // Битовая маска для расшифровки
END_VAR
VAR
	stError : ST_ROBOT_ERROR; // Представление ошибок отдельными флагами
END_VAR
stError.WRONG_ACTION := (dwError AND ERR_ROBOT_WRONG_ACTION) <> DWORD#0;
stError.MOTION_ERROR := (dwError AND ERR_ROBOT_MOTION) <> DWORD#0;
stError.GRIPPER_ERROR := (dwError AND ERR_ROBOT_GRIPPER) <> DWORD#0;
stError.MODBUS_COMMUNICATION_ERROR := (dwError AND ERR_ROBOT_MODBUS_COMM) <> DWORD#0;
stError.EXTERNAL_ROBOT_ALARM := (dwError AND ERR_EXTERNAL_ROBOT) <> DWORD#0;
stError.MODBUS_ERROR := stError.MODBUS_COMMUNICATION_ERROR OR stError.EXTERNAL_ROBOT_ALARM;
stError.STOP_ERROR := (dwError AND ERR_ROBOT_STOP) <> DWORD#0;

UpdateErrorView := stError;
END_METHOD

END_FUNCTION_BLOCK

// Device/Application/FB/FB_MAGAZINE
FUNCTION_BLOCK FB_MAGAZINE
VAR_INPUT
	xIoManual : BOOL; // Передача выходов оператору отменяет пошаговую операцию
	uiMagazineId : UINT; // Идентификатор экземпляра 1..2
	xPointsConfigured : BOOL; // Настроена база этого магазина с Safe Z и Change Z
	xMechanismReady : BOOL := TRUE;
	xInventoryChanged : BOOL; // Сменился рабочий банк или оператор изменил его содержимое
	xTestInitialize : BOOL;
	xTestEnabled : BOOL;
	stRobotStatus     : ST_ROBOT_STATUS; // Текущие статусы робота
	astMachineStatus  : ARRAY [1..3] OF ST_MACHINE_PUBLIC; // Статусы станков для определения оставшейся работы
	auiMachineType    : ARRAY [1..3] OF UINT; // Тип детали, закреплённый за каждым станком
	stMagazineCommand : ST_MAGAZINE_COMMAND; // Команда магазина от автоматической логики
	stHmiCommand      : ST_ROBOT_COMMAND; // Ручная команда магазина с HMI
	xManual           : BOOL; // Разрешение ручного управления
	xReset            : BOOL; // Сброс ошибок магазина
	xGlobalError      : BOOL; // Глобальная ошибка ячейки
	xHmiEnable        : BOOL; // Импульс включения магазина с HMI
	xHmiDisable       : BOOL; // Импульс отключения магазина с HMI
	xHmiFillBlanks    : BOOL; // Заполнить все активные слоты матрицы заготовками
	xHmiClear         : BOOL; // Полностью очистить содержимое магазина
	xHmiCycleSlot     : BOOL; // Переключить содержимое выбранного слота
	xHmiApplySlot     : BOOL; // Явно записать состояние и тип выбранного слота
	xHmiApplyPitchX   : BOOL; // Применить новый общий шаг слотов по X
	xHmiApplyPitchY   : BOOL; // Применить новый общий шаг слотов по Y
	uiHmiEditSlot     : UINT; // Номер слота для ручного редактирования
	uiHmiEditDetailType : UINT; // 0=NONE, 1=BLANK, 2=DETAIL
	uiHmiEditProductType : UINT; // Тип изделия 1..3
	lrHmiEditPitchX   : LREAL;
	lrHmiEditPitchY   : LREAL;
	xRobotOwnsMagazine : BOOL; // Автомат удерживает этот магазин в текущем цикле
	xRobotCanWorkWithMagazine : BOOL; // Интерфейс и точки готовы для роботной операции, не для включения магазина
	xSharedGeometryEditAllowed : BOOL; // Оба магазина выключены; общий шаг можно менять
	uiRows            : UINT; // Число строк матрицы магазина
	uiColumns         : UINT; // Число столбцов матрицы магазина
	uiTypeCount       : UINT; // Количество настроенных типов заготовок, 1..3
	auiSlotType       : ARRAY [1..GVL_CELL_SETTINGS.NumberDetail] OF UINT; // Тип секции каждого слота
	FaultRequest  : ST_MAGAZINE_FAULT_REQUEST; // Единый контракт диагностической инъекции
END_VAR
VAR_OUTPUT
	Command : ST_ROBOT_COMMAND; // Текущая пошаговая команда роботу
	Status  : ST_MAGAZINE_STATUS; // Рабочие статусы магазина
	Diag    : ST_MAGAZINE_DIAG; // Состояние автомата магазина
	Error   : ST_MAGAZINE_ERRORS; // Активные и последние ошибки
	FaultStatus : ST_FAULT_INJECTION_STATUS; // Состояние инжектора для HMI
END_VAR
VAR_IN_OUT
	stInventory : ST_MAGAZINE_INVENTORY; // Единственная кассета текущего магазина
	lrPitchX : LREAL; // Общий фактический шаг слотов по X
	lrPitchY : LREAL; // Общий фактический шаг слотов по Y
END_VAR
VAR
	eGrantedOperation : E_MAGAZINE_OPERATION; // Доступная операция магазина
	eActualOperation  : E_MAGAZINE_OPERATION; // Выполняемая операция магазина

	rtExecute          : R_TRIG; // Фронт команды запуска
	rtEnable           : R_TRIG; // Фронт команды включения
	rtDisable          : R_TRIG; // Фронт команды отключения
	rtFillBlanks       : R_TRIG; // Фронт заполнения магазина заготовками
	rtClear            : R_TRIG; // Фронт очистки магазина
	rtCycleSlot        : R_TRIG; // Фронт изменения выбранного слота
	rtApplySlot        : R_TRIG; // Фронт явной записи выбранного слота
	rtApplyPitchX      : R_TRIG;
	rtApplyPitchY      : R_TRIG;
	rtReset            : R_TRIG; // Фронт команды сброса магазина

	xExecuteRequest    : BOOL; // Активный запрос выполнения операции
	xResetRequest      : BOOL; // Активный запрос сброса
	xStopRequest       : BOOL; // Активный запрос остановки
	xManualCommand     : BOOL; // Команда получена из ручного интерфейса
	xDisableRequest    : BOOL; // Сохранённый запрос отключения после текущей операции
	xRobotInMagazineContext : BOOL; // Робот находится в рабочей зоне магазина
	xFaultContextCaptured : BOOL; // Контекст робота зафиксирован при входе в ERROR
	xRobotInMagazineAtFault : BOOL; // Робот был в рабочей зоне этого магазина при ошибке
	xRobotStopRequired : BOOL; // Итоговая реакция ROBOT_STOP, сформированная магазином
	xRobotResetDependencyReady : BOOL; // Каскадная ошибка робота может быть сброшена тем же импульсом

	iActiveSlotCount   : SINT; // Число активных слотов выбранной матрицы
	iInventoryIndex    : SINT; // Индекс изменения содержимого магазина
	iTakeSlot          : SINT; // Слот выбранной заготовки
	iPutSlot           : SINT; // Выбранный свободный слот
	iActiveSlot        : SINT; // Единственный слот текущего элементарного движения
	xInventoryCommitted: BOOL; // Все изменения слотов текущей операции подтверждены
	xTakeSlotCommitted  : BOOL; // Изъятие заготовки отражено в матрице после закрытия захвата
	xPutSlotCommitted   : BOOL; // Укладка груза отражена в матрице после открытия захвата
	xRobotCommandStarted : BOOL; // Текущий элементарный шаг действительно принят FB_ROBOT
	xOperationSequenceComplete : BOOL; // Все шаги операции подтверждены до изменения матрицы
	xTakeSlotValid     : BOOL; // Проверка диапазона до обращения к массиву слотов
	xPutSlotValid      : BOOL;
	xTakeSlotHasBlank  : BOOL;
	xPutSlotEmpty      : BOOL;
	xChangeTakeFirst   : BOOL; // CHANGE в одном слоте: сначала TAKE, затем PUT
	xPutProductTypeValid : BOOL;
	uiStep             : UINT; // Шаг последовательности робота
	uiIndex            : UINT; // Индекс слота для расчёта координат

	stActiveRobotCommand : ST_ROBOT_COMMAND; // Команда роботу текущего шага
	xFinishedCondition   : BOOL; // Текущее содержимое не позволяет продолжить цикл
	xFinishedLatched     : BOOL; // Завершение этой палеты не отменяется работой другого магазина
	xMachineHasRelevantPart : BOOL; // В доступном станке есть заготовка, обработка или готовая деталь
	xMachineHasDestination : BOOL; // Для оставшейся работы есть свободный слот соответствующего типа
	xAllSlotsDetails    : BOOL; // Все активные слоты заполнены готовыми деталями
	xNoBlankNoMachinePart : BOOL; // Нет заготовок и нет доступной работы в станках
	xNoBlankNoDestination : BOOL; // Нет заготовок и нет места для возврата груза
	uiMachineIndex      : UINT; // Индекс станка при расчёте завершения магазина
	uiMachineTypeIndex  : UINT; // Тип детали проверяемого станка
	uiPutProductType    : UINT; // Тип груза, защёлкнутый до физического PUT
	fbFaultInjector      : FB_MAGAZINE_FAULT_INJECTOR; // Безопасный сценарий ошибки до движения
	xFaultAllowed        : BOOL; // Владелец разрешает синтетическую проверку
	xStartupInitialized  : BOOL;
	udiProducedPartsTotal : UDINT; // Монотонный счётчик подтверждённых укладок готовых деталей
END_VAR
VAR CONSTANT
	ERR_WRONG_OPERATION : DWORD := DWORD#16#0000_0001; // Недопустимая операция магазина
	ERR_NO_BLANK        : DWORD := DWORD#16#0000_0002; // В магазине нет заготовки
	ERR_NO_FREE_SLOT    : DWORD := DWORD#16#0000_0004; // В магазине нет свободного слота
	ERR_INVALID_SLOT    : DWORD := DWORD#16#0000_0008; // Недопустимый номер слота
	ERR_SLOT_CONTENT    : DWORD := DWORD#16#0000_0010; // Содержимое слота не соответствует операции
	ERR_ROBOT           : DWORD := DWORD#16#0000_0020; // Ошибка робота при операции магазина
	ERR_GLOBAL_STOP     : DWORD := DWORD#16#0000_0040; // Остановка по глобальной ошибке
	ERR_GEOMETRY        : DWORD := DWORD#16#0000_0080; // Ошибка параметров матрицы магазина
	MASK_EQUIPMENT_ERROR : DWORD := ERR_WRONG_OPERATION OR ERR_NO_BLANK
		OR ERR_NO_FREE_SLOT OR ERR_INVALID_SLOT OR ERR_SLOT_CONTENT OR ERR_GEOMETRY;
	WRN_RESET_EXECUTE_ACTIVE : UINT := 1; // Операция магазина ещё активна
	WRN_RESET_GLOBAL_ERROR   : UINT := 2; // Глобальная ошибка ещё активна
	WRN_RESET_ROBOT_ERROR    : UINT := 3; // Ошибка робота ещё активна
	WRN_ENABLE_GLOBAL_ERROR  : UINT := 4; // Включение запрещено глобальной ошибкой
	WRN_ENABLE_CONTENT       : UINT := 5; // Архив: содержимое больше не блокирует включение
	WRN_DISABLE_PENDING      : UINT := 6; // Отключение магазина уже запрошено
	WRN_FILL_ENABLED         : UINT := 7; // Заполнение запрещено для включённого магазина
	WRN_FILL_GEOMETRY        : UINT := 8; // Активная матрица магазина задана неверно
	WRN_CLEAR_ENABLED        : UINT := 9; // Очистка запрещена для включённого магазина
	WRN_SIM_ERROR_NOT_ALLOWED: UINT := 10; // Тестовая ошибка запрещена текущим состоянием
	WRN_EDIT_REJECTED : UINT := 14; // Редактирование включённого/занятого магазина запрещено
	WRN_GEOMETRY_EDIT_REJECTED : UINT := 16; // PLC отклонил изменение общего шага X/Y
	WRN_ENABLE_GEOMETRY      : UINT := 15; // Геометрия магазина не позволяет включение
	WRN_ENABLE_OWN_ERROR     : UINT := 17; // Включение запрещено собственной ошибкой магазина
	WRN_ENABLE_POINTS        : UINT := 18; // Не настроена база этого магазина или её Z-смещения
END_VAR

// Инвентарь загружает владелец банков RunTwoPallet; здесь сбрасывается только автомат.
IF NOT xStartupInitialized THEN
	xFinishedLatched := FALSE;
	xFaultContextCaptured := FALSE;
	xRobotInMagazineAtFault := FALSE;
	xRobotStopRequired := FALSE;
	xStartupInitialized := TRUE;
END_IF;

IF xTestInitialize THEN
	xFinishedLatched := FALSE;
	IF xTestEnabled AND xPointsConfigured THEN
		Diag.eState := E_MAGAZINE_STATE.IDLE;
	ELSE
		Diag.eState := E_MAGAZINE_STATE.DISABLED;
	END_IF;
	Error.dwErrorActive := DWORD#0;
	Error.dwAlarmActive := DWORD#0;
	eGrantedOperation := E_MAGAZINE_OPERATION.NONE;
	eActualOperation := E_MAGAZINE_OPERATION.NONE;
	xExecuteRequest := FALSE;
	xResetRequest := FALSE;
	xStopRequest := FALSE;
	xManualCommand := FALSE;
	xDisableRequest := FALSE;
	iTakeSlot := SINT#0;
	iPutSlot := SINT#0;
	xChangeTakeFirst := FALSE;
	iActiveSlot := SINT#0;
	xInventoryCommitted := FALSE;
	xTakeSlotCommitted := FALSE;
	xPutSlotCommitted := FALSE;
	xRobotCommandStarted := FALSE;
	xOperationSequenceComplete := FALSE;
	xFaultContextCaptured := FALSE;
	xRobotInMagazineAtFault := FALSE;
	xRobotStopRequired := FALSE;
	uiStep := UINT#0;
	stActiveRobotCommand.xExecute := FALSE;
	stActiveRobotCommand.xStop := FALSE;
	stActiveRobotCommand.xReset := FALSE;
	stActiveRobotCommand.eAction := E_ROBOT_ACTION.NONE;
	stActiveRobotCommand.eSetPoint := E_POINT_NAME.NONE;
	stActiveRobotCommand.iActiveSlot := SINT#0;
	stActiveRobotCommand.uiMagazineId := uiMagazineId;
END_IF;

IF xInventoryChanged THEN
	xFinishedLatched := FALSE;
END_IF;

rtFillBlanks(CLK := xHmiFillBlanks);
rtClear(CLK := xHmiClear);
rtCycleSlot(CLK := xHmiCycleSlot);
rtApplySlot(CLK := xHmiApplySlot);
rtApplyPitchX(CLK := xHmiApplyPitchX);
rtApplyPitchY(CLK := xHmiApplyPitchY);

IF (uiRows > UINT#0)
AND (uiColumns > UINT#0)
AND ((uiRows * uiColumns) <= SINT_TO_UINT(GVL_CELL_SETTINGS.MagazineSlots)) THEN
	iActiveSlotCount := UINT_TO_SINT(uiRows * uiColumns);
ELSE
	iActiveSlotCount := SINT#0;
END_IF;

// Ручная роботная команда принадлежит только выбранному магазину.
xManualCommand := xManual
	AND (
		(stHmiCommand.eSetPoint = E_POINT_NAME.MAGAZINE_TAKE_DETAIL)
		OR (stHmiCommand.eSetPoint = E_POINT_NAME.MAGAZINE_PUT_DETAIL)
		OR (stHmiCommand.eSetPoint = E_POINT_NAME.MAGAZINE_CHANGE_DETAIL)
		OR (stHmiCommand.eSetPoint = E_POINT_NAME.MAGAZINE_RETURN_BLANK)
	)
	AND ((stHmiCommand.uiMagazineId = uiMagazineId)
		OR ((stHmiCommand.uiMagazineId = UINT#0) AND (uiMagazineId = UINT#1)));

IF xManual THEN
	IF xManualCommand THEN
		xExecuteRequest := stHmiCommand.xExecute;
		xStopRequest := stHmiCommand.xStop;
	ELSE
		xExecuteRequest := FALSE;
		xStopRequest := FALSE;
	END_IF;
ELSE
	xExecuteRequest := stMagazineCommand.xExecute;
	xStopRequest := stMagazineCommand.xStop;
END_IF;

// Контекст запрещает редактирование и завершает отложенное отключение только
// после фактического выхода робота из конкретного магазина.
xRobotInMagazineContext := (stRobotStatus.uiMagazineContext = uiMagazineId)
	OR ((stRobotStatus.uiMagazineContext = UINT#0)
		AND (xRobotOwnsMagazine OR xManualCommand)
		AND ((stRobotStatus.eCurrentPoint = E_POINT_NAME.MAGAZINE_IN_SLOT)
			OR (stRobotStatus.eCurrentPoint = E_POINT_NAME.MAGAZINE_CHANGE)));
xRobotInMagazineContext := xRobotInMagazineContext
	OR ((xRobotOwnsMagazine OR xManualCommand)
		AND (Diag.eState = E_MAGAZINE_STATE.ROBOT_COMMAND)
		AND (stActiveRobotCommand.eAction = E_ROBOT_ACTION.MOVE_TO_POINT)
		AND ((stActiveRobotCommand.eSetPoint = E_POINT_NAME.MAGAZINE_IN_SLOT)
			OR (stActiveRobotCommand.eSetPoint = E_POINT_NAME.MAGAZINE_CHANGE)));

// Единственную кассету можно менять только у технологически выключенного
// магазина, когда робот не находится внутри и не владеет текущей операцией.
Status.xEditAllowed := ((Diag.eState = E_MAGAZINE_STATE.DISABLED)
		OR (Diag.eState = E_MAGAZINE_STATE.ERROR))
	AND NOT xRobotOwnsMagazine
	AND NOT xRobotInMagazineContext
	AND NOT xGlobalError;
Status.xPitchEditAllowed := Status.xEditAllowed AND xSharedGeometryEditAllowed;

// Шаг матрицы общий для двух магазинов, поэтому менять его разрешено только
// когда оба магазина выключены. Смещения Z принадлежат базовым точкам магазина.
IF rtApplyPitchX.Q
AND Status.xEditAllowed
AND xSharedGeometryEditAllowed
AND (lrHmiEditPitchX >= LREAL#1.0)
AND (lrHmiEditPitchX <= LREAL#5000.0) THEN
	lrPitchX := lrHmiEditPitchX;
END_IF;
IF rtApplyPitchY.Q
AND Status.xEditAllowed
AND xSharedGeometryEditAllowed
AND (lrHmiEditPitchY >= LREAL#1.0)
AND (lrHmiEditPitchY <= LREAL#5000.0) THEN
	lrPitchY := lrHmiEditPitchY;
END_IF;
IF rtClear.Q AND Status.xEditAllowed THEN
	xFinishedLatched := FALSE;
	FOR iInventoryIndex := 1 TO GVL_CELL_SETTINGS.MagazineSlots DO
		stInventory.aSlots[iInventoryIndex].xInPosition := FALSE;
		stInventory.aSlots[iInventoryIndex].eDetailType := E_DETAIL_TYPE.NONE;
		stInventory.aSlots[iInventoryIndex].uiProductType := UINT#0;
	END_FOR;
ELSIF rtFillBlanks.Q
AND (iActiveSlotCount > SINT#0)
AND Status.xEditAllowed THEN
	xFinishedLatched := FALSE;
	FOR iInventoryIndex := 1 TO GVL_CELL_SETTINGS.MagazineSlots DO
		stInventory.aSlots[iInventoryIndex].xInPosition := iInventoryIndex <= iActiveSlotCount;
		IF iInventoryIndex <= iActiveSlotCount THEN
			stInventory.aSlots[iInventoryIndex].eDetailType := E_DETAIL_TYPE.BLANK;
			stInventory.aSlots[iInventoryIndex].uiProductType := auiSlotType[iInventoryIndex];
		ELSE
			stInventory.aSlots[iInventoryIndex].eDetailType := E_DETAIL_TYPE.NONE;
			stInventory.aSlots[iInventoryIndex].uiProductType := UINT#0;
		END_IF;
	END_FOR;
ELSIF rtApplySlot.Q
AND Status.xEditAllowed
AND (uiHmiEditSlot >= UINT#1)
AND (uiHmiEditSlot <= SINT_TO_UINT(iActiveSlotCount))
AND (uiHmiEditDetailType <= UINT#2)
AND ((uiHmiEditDetailType = UINT#0)
	OR ((uiHmiEditProductType >= UINT#1) AND (uiHmiEditProductType <= uiTypeCount))) THEN
	xFinishedLatched := FALSE;
	iInventoryIndex := UINT_TO_SINT(uiHmiEditSlot);
	CASE uiHmiEditDetailType OF
		UINT#0:
			stInventory.aSlots[iInventoryIndex].xInPosition := FALSE;
			stInventory.aSlots[iInventoryIndex].eDetailType := E_DETAIL_TYPE.NONE;
			stInventory.aSlots[iInventoryIndex].uiProductType := UINT#0;
		UINT#1:
			stInventory.aSlots[iInventoryIndex].xInPosition := TRUE;
			stInventory.aSlots[iInventoryIndex].eDetailType := E_DETAIL_TYPE.BLANK;
			stInventory.aSlots[iInventoryIndex].uiProductType := uiHmiEditProductType;
		UINT#2:
			stInventory.aSlots[iInventoryIndex].xInPosition := TRUE;
			stInventory.aSlots[iInventoryIndex].eDetailType := E_DETAIL_TYPE.DETAIL;
			stInventory.aSlots[iInventoryIndex].uiProductType := uiHmiEditProductType;
	END_CASE;
ELSIF rtCycleSlot.Q
AND Status.xEditAllowed
AND (uiHmiEditSlot >= UINT#1)
AND (uiHmiEditSlot <= SINT_TO_UINT(iActiveSlotCount)) THEN
	xFinishedLatched := FALSE;
	iInventoryIndex := UINT_TO_SINT(uiHmiEditSlot);
	IF NOT stInventory.aSlots[iInventoryIndex].xInPosition
	OR (stInventory.aSlots[iInventoryIndex].eDetailType = E_DETAIL_TYPE.NONE) THEN
		stInventory.aSlots[iInventoryIndex].xInPosition := TRUE;
		stInventory.aSlots[iInventoryIndex].eDetailType := E_DETAIL_TYPE.BLANK;
		stInventory.aSlots[iInventoryIndex].uiProductType := auiSlotType[iInventoryIndex];
	ELSE
		stInventory.aSlots[iInventoryIndex].xInPosition := FALSE;
		stInventory.aSlots[iInventoryIndex].eDetailType := E_DETAIL_TYPE.NONE;
		stInventory.aSlots[iInventoryIndex].uiProductType := UINT#0;
	END_IF;
END_IF;

// При смене банка проверка завершения использует его текущую карту типов,
// а не свободные слоты прежней палеты с прошлого скана.
UpdateTypeStatus(stMagazineInventory := stInventory);

IF iActiveSlotCount > SINT#0 THEN
	Status.iCurrentBlank := FindBlank(stDetail := stInventory.aSlots, iSlotCount := iActiveSlotCount);
	Status.iCurrentFreeSlot := FindFreeSlot(stDetail := stInventory.aSlots, iSlotCount := iActiveSlotCount);
ELSE
	Status.iCurrentBlank := SINT#0;
	Status.iCurrentFreeSlot := SINT#0;
END_IF;

Status.xOutBlank := Status.iCurrentBlank = SINT#0;
Status.xOutFreeSlot := Status.iCurrentFreeSlot = SINT#0;
Status.xCanTake := NOT Status.xOutBlank;
Status.xCanPut := NOT Status.xOutFreeSlot;
Status.xCanChange := Status.xCanTake; // Изъятие заготовки само освобождает место
Status.xCanEnable := FALSE;

// Для PUT/возврата заготовки нужен пустой слот. Готовую деталь можно обменять
// на заготовку в одном занятом слоте, если первый захват свободен и открыт.
IF stRobotStatus.xBlankAvailable OR stRobotStatus.xDetailAvailable THEN
	Status.xCanEnable := Status.xCanPut;
ELSIF NOT stRobotStatus.xBlankAvailable AND NOT stRobotStatus.xDetailAvailable THEN
	Status.xCanEnable := Status.xCanTake;
END_IF;

IF stRobotStatus.xDetailAvailable AND NOT stRobotStatus.xBlankAvailable
AND stRobotStatus.xGripper1Open AND Status.xCanChange THEN
	Status.xCanEnable := TRUE;
END_IF;

// Отсутствие заготовок не завершает магазин, пока из станков ещё можно вернуть
// готовую деталь в свободный слот соответствующего типа.
xMachineHasRelevantPart := FALSE;
xMachineHasDestination := FALSE;
FOR uiMachineIndex := UINT#1 TO UINT#3 DO
	IF astMachineStatus[uiMachineIndex].xEnabled
	AND NOT astMachineStatus[uiMachineIndex].xError
	AND (astMachineStatus[uiMachineIndex].xProcessing
		OR ((astMachineStatus[uiMachineIndex].ePartState = E_PART_STATE.LOADED)
			AND ((astMachineStatus[uiMachineIndex].ePartType = E_PART_TYPE.PART)
				OR (astMachineStatus[uiMachineIndex].ePartType = E_PART_TYPE.DETAIL)))) THEN
		xMachineHasRelevantPart := TRUE;
		uiMachineTypeIndex := auiMachineType[uiMachineIndex];
		IF (uiMachineTypeIndex >= UINT#1)
		AND (uiMachineTypeIndex <= UINT#3)
		AND (Status.stTypeStatus.aiFreeSlot[uiMachineTypeIndex] > SINT#0) THEN
			xMachineHasDestination := TRUE;
		END_IF;
	END_IF;
END_FOR;

IF NOT stRobotStatus.xBlankAvailable
AND NOT stRobotStatus.xDetailAvailable
AND xMachineHasDestination THEN
	Status.xCanEnable := TRUE;
END_IF;

Status.xEnableCheckRobotReady := xRobotCanWorkWithMagazine AND xMechanismReady;
Status.xEnableCheckRobotReleased := NOT xRobotInMagazineContext;
Status.xEnableCheckNoError := NOT xGlobalError
	AND (Diag.eState <> E_MAGAZINE_STATE.ERROR)
	AND (Error.dwErrorActive = DWORD#0);
Status.xEnableCheckContent := Status.xCanEnable;
Status.xEnableCheckGeometry := (iActiveSlotCount > SINT#0)
	AND (lrPitchX >= LREAL#1.0)
	AND (lrPitchX <= LREAL#5000.0)
	AND (lrPitchY >= LREAL#1.0)
	AND (lrPitchY <= LREAL#5000.0);
// Включение требует собственную базовую точку магазина. Готовность интерфейса,
// положение робота и содержимое палеты проверяются при роботной операции.
Status.xEnableSequenceAllowed := (Diag.eState = E_MAGAZINE_STATE.DISABLED)
	AND Status.xEnableCheckNoError
	AND Status.xEnableCheckGeometry
	AND xPointsConfigured;

// Finished остаётся прежним по смыслу, но теперь оценивает единственную кассету.
xAllSlotsDetails := iActiveSlotCount > SINT#0;
IF xAllSlotsDetails THEN
	FOR uiIndex := UINT#1 TO SINT_TO_UINT(iActiveSlotCount) DO
		IF NOT stInventory.aSlots[UINT_TO_SINT(uiIndex)].xInPosition
		OR (stInventory.aSlots[UINT_TO_SINT(uiIndex)].eDetailType <> E_DETAIL_TYPE.DETAIL) THEN
			xAllSlotsDetails := FALSE;
		END_IF;
	END_FOR;
END_IF;
xNoBlankNoMachinePart := Status.xOutBlank AND NOT xMachineHasRelevantPart;
xNoBlankNoDestination := Status.xOutBlank AND NOT xMachineHasDestination;
xFinishedCondition :=
	(NOT stRobotStatus.xBlankAvailable AND NOT stRobotStatus.xDetailAvailable)
	AND (xAllSlotsDetails OR xNoBlankNoMachinePart OR xNoBlankNoDestination);

eGrantedOperation := E_MAGAZINE_OPERATION.NONE;
IF stRobotStatus.xBlankAvailable
AND stRobotStatus.xDetailAvailable
AND Status.xCanPut THEN
	// Сначала освобождается захват готовой детали; заготовка остаётся у робота.
	eGrantedOperation := E_MAGAZINE_OPERATION.PUT;
ELSIF NOT Status.xOutBlank
AND NOT stRobotStatus.xBlankAvailable
AND NOT stRobotStatus.xDetailAvailable THEN
	eGrantedOperation := E_MAGAZINE_OPERATION.TAKE;
ELSIF NOT Status.xOutBlank
AND stRobotStatus.xGripper1Open
AND NOT stRobotStatus.xBlankAvailable
AND stRobotStatus.xDetailAvailable THEN
	eGrantedOperation := E_MAGAZINE_OPERATION.CHANGE;
ELSIF NOT Status.xOutFreeSlot
AND stRobotStatus.xDetailAvailable THEN
	eGrantedOperation := E_MAGAZINE_OPERATION.PUT;
END_IF;

xResetRequest := xReset;
rtReset(CLK := xResetRequest);

xRobotResetDependencyReady := (((Error.dwErrorActive AND ERR_ROBOT) = DWORD#0)
		AND NOT xRobotInMagazineAtFault)
	OR NOT stRobotStatus.xError
	OR stRobotStatus.xResetAllowed;

IF rtReset.Q
AND (Diag.eState = E_MAGAZINE_STATE.ERROR) THEN
	IF xExecuteRequest THEN
		Diag.stWarning.uiCode := WRN_RESET_EXECUTE_ACTIVE;
	ELSIF xGlobalError THEN
		Diag.stWarning.uiCode := WRN_RESET_GLOBAL_ERROR;
	ELSIF stRobotStatus.xError
	AND NOT stRobotStatus.xResetAllowed THEN
		Diag.stWarning.uiCode := WRN_RESET_ROBOT_ERROR;
	ELSE
		Diag.stWarning.uiCode := UINT#0;
	END_IF;

	IF Diag.stWarning.uiCode <> UINT#0 THEN
		Diag.stWarning.udiSequence := Diag.stWarning.udiSequence + UDINT#1;
		IF Diag.stWarning.udiSequence = UDINT#0 THEN
			Diag.stWarning.udiSequence := UDINT#1;
		END_IF;
	END_IF;
END_IF;

rtEnable(CLK := xHmiEnable OR (NOT xManual AND stMagazineCommand.xEnable));
rtDisable(CLK := xHmiDisable OR (NOT xManual AND stMagazineCommand.xDisable));

IF rtEnable.Q
AND (Diag.eState = E_MAGAZINE_STATE.DISABLED)
AND NOT Status.xEnableSequenceAllowed THEN
	IF NOT xPointsConfigured THEN
		Diag.stWarning.uiCode := WRN_ENABLE_POINTS;
	ELSIF xGlobalError THEN
		Diag.stWarning.uiCode := WRN_ENABLE_GLOBAL_ERROR;
	ELSIF NOT Status.xEnableCheckGeometry THEN
		Diag.stWarning.uiCode := WRN_ENABLE_GEOMETRY;
	ELSE
		Diag.stWarning.uiCode := WRN_ENABLE_OWN_ERROR;
	END_IF;
	Diag.stWarning.udiSequence := Diag.stWarning.udiSequence + UDINT#1;
	IF Diag.stWarning.udiSequence = UDINT#0 THEN
		Diag.stWarning.udiSequence := UDINT#1;
	END_IF;
ELSIF rtDisable.Q
AND xHmiDisable
AND xDisableRequest THEN
	Diag.stWarning.uiCode := WRN_DISABLE_PENDING;
	Diag.stWarning.udiSequence := Diag.stWarning.udiSequence + UDINT#1;
	IF Diag.stWarning.udiSequence = UDINT#0 THEN
		Diag.stWarning.udiSequence := UDINT#1;
	END_IF;
ELSIF rtFillBlanks.Q
AND (iActiveSlotCount = 0) THEN
	Diag.stWarning.uiCode := WRN_FILL_GEOMETRY;
	Diag.stWarning.udiSequence := Diag.stWarning.udiSequence + UDINT#1;
	IF Diag.stWarning.udiSequence = UDINT#0 THEN
		Diag.stWarning.udiSequence := UDINT#1;
	END_IF;
ELSIF rtFillBlanks.Q
AND NOT Status.xEditAllowed THEN
	Diag.stWarning.uiCode := WRN_FILL_ENABLED;
	Diag.stWarning.udiSequence := Diag.stWarning.udiSequence + UDINT#1;
	IF Diag.stWarning.udiSequence = UDINT#0 THEN
		Diag.stWarning.udiSequence := UDINT#1;
	END_IF;
ELSIF rtClear.Q
AND NOT Status.xEditAllowed THEN
	Diag.stWarning.uiCode := WRN_CLEAR_ENABLED;
	Diag.stWarning.udiSequence := Diag.stWarning.udiSequence + UDINT#1;
	IF Diag.stWarning.udiSequence = UDINT#0 THEN
		Diag.stWarning.udiSequence := UDINT#1;
	END_IF;
ELSIF (rtApplyPitchX.Q
	AND (NOT Status.xEditAllowed
		OR NOT xSharedGeometryEditAllowed
		OR (lrHmiEditPitchX < LREAL#1.0)
		OR (lrHmiEditPitchX > LREAL#5000.0)))
OR (rtApplyPitchY.Q
	AND (NOT Status.xEditAllowed
		OR NOT xSharedGeometryEditAllowed
		OR (lrHmiEditPitchY < LREAL#1.0)
		OR (lrHmiEditPitchY > LREAL#5000.0))) THEN
	Diag.stWarning.uiCode := WRN_GEOMETRY_EDIT_REJECTED;
	Diag.stWarning.udiSequence := Diag.stWarning.udiSequence + UDINT#1;
	IF Diag.stWarning.udiSequence = UDINT#0 THEN
		Diag.stWarning.udiSequence := UDINT#1;
	END_IF;
ELSIF rtApplySlot.Q
AND ((uiHmiEditSlot < UINT#1)
	OR (uiHmiEditSlot > SINT_TO_UINT(iActiveSlotCount))
	OR (uiHmiEditDetailType > UINT#2)
	OR ((uiHmiEditDetailType <> UINT#0)
		AND ((uiHmiEditProductType < UINT#1) OR (uiHmiEditProductType > uiTypeCount)))
	OR NOT Status.xEditAllowed) THEN
	Diag.stWarning.uiCode := WRN_EDIT_REJECTED;
	Diag.stWarning.udiSequence := Diag.stWarning.udiSequence + UDINT#1;
	IF Diag.stWarning.udiSequence = UDINT#0 THEN
		Diag.stWarning.udiSequence := UDINT#1;
	END_IF;
ELSIF rtCycleSlot.Q
AND ((uiHmiEditSlot < UINT#1)
	OR (uiHmiEditSlot > SINT_TO_UINT(iActiveSlotCount))
	OR NOT Status.xEditAllowed) THEN
	Diag.stWarning.uiCode := WRN_EDIT_REJECTED;
	Diag.stWarning.udiSequence := Diag.stWarning.udiSequence + UDINT#1;
	IF Diag.stWarning.udiSequence = UDINT#0 THEN
		Diag.stWarning.udiSequence := UDINT#1;
	END_IF;
END_IF;

IF rtDisable.Q THEN
	xDisableRequest := TRUE;
END_IF;

rtExecute(CLK := xExecuteRequest);

// Синтетический сценарий входит только в проверочный шаг CHOOSE и не выдаёт
// команду движения роботу до формирования выбранной штатной ошибки.
xFaultAllowed := ((Diag.eState = E_MAGAZINE_STATE.DISABLED)
	OR (Diag.eState = E_MAGAZINE_STATE.IDLE))
	AND NOT xExecuteRequest
	AND NOT xGlobalError
	AND NOT stRobotStatus.xBusy
	AND NOT stRobotStatus.xError
	AND (Error.dwErrorActive = DWORD#0);

fbFaultInjector(
	Request := FaultRequest,
	xOwnerAllowed := xFaultAllowed,
	xComplete := Diag.eState = E_MAGAZINE_STATE.ERROR
);
FaultStatus := fbFaultInjector.Status;

IF fbFaultInjector.Status.xRejected THEN
	Diag.stWarning.uiCode := WRN_SIM_ERROR_NOT_ALLOWED;
	Diag.stWarning.udiSequence := Diag.stWarning.udiSequence + UDINT#1;
	IF Diag.stWarning.udiSequence = UDINT#0 THEN
		Diag.stWarning.udiSequence := UDINT#1;
	END_IF;
END_IF;

// Значения команды роботу по умолчанию.
Command.xExecute := FALSE;
Command.xStop := FALSE;
Command.xReset := xResetRequest;
Command.eAction := E_ROBOT_ACTION.NONE;
Command.eSetPoint := E_POINT_NAME.NONE;
Command.iActiveSlot := 0;
Command.uiMagazineId := UINT#0;

// Ошибка робота в рабочей зоне принадлежит одновременно роботу и магазину.
IF xRobotInMagazineContext
AND stRobotStatus.xError
AND (Diag.eState <> E_MAGAZINE_STATE.ERROR) THEN
	Error.dwErrorActive := Error.dwErrorActive OR ERR_ROBOT;
	Diag.eState := E_MAGAZINE_STATE.ERROR;
END_IF;

IF xGlobalError
AND (Diag.eState <> E_MAGAZINE_STATE.DISABLED)
AND (Diag.eState <> E_MAGAZINE_STATE.IDLE)
AND (Diag.eState <> E_MAGAZINE_STATE.ERROR) THEN
	Error.dwErrorActive := Error.dwErrorActive OR ERR_GLOBAL_STOP;
	Diag.eState := E_MAGAZINE_STATE.ERROR;
END_IF;

// Сохраняем уже подтверждённые изменения слотов и первичную аварию,
// но не оставляем команду, которая продолжится после возврата I/O программе.
IF xIoManual THEN
	xExecuteRequest := FALSE;
	xStopRequest := FALSE;
	xDisableRequest := FALSE;
	xRobotCommandStarted := FALSE;
	xOperationSequenceComplete := FALSE;
	eActualOperation := E_MAGAZINE_OPERATION.NONE;
	stActiveRobotCommand.xExecute := FALSE;
	IF Diag.eState <> E_MAGAZINE_STATE.ERROR THEN
		Diag.eState := E_MAGAZINE_STATE.DISABLED;
	END_IF;
END_IF;

CASE Diag.eState OF
	E_MAGAZINE_STATE.DISABLED:
		xDisableRequest := FALSE;
		IF fbFaultInjector.Status.xBusy THEN
			iTakeSlot := 1;
			iPutSlot := 1;
			IF fbFaultInjector.xWrongOperation THEN
				eActualOperation := E_MAGAZINE_OPERATION.NONE;
			ELSIF fbFaultInjector.xNoFreeSlot THEN
				eActualOperation := E_MAGAZINE_OPERATION.PUT;
			ELSE
				eActualOperation := E_MAGAZINE_OPERATION.TAKE;
			END_IF;
			Diag.eState := E_MAGAZINE_STATE.CHOOSE;
		ELSIF rtEnable.Q AND NOT xIoManual
		AND Status.xEnableSequenceAllowed THEN
			Diag.eState := E_MAGAZINE_STATE.IDLE;
		END_IF;

	E_MAGAZINE_STATE.IDLE:
		uiStep := 0;
		eActualOperation := E_MAGAZINE_OPERATION.NONE;
		xInventoryCommitted := FALSE;
		xTakeSlotCommitted := FALSE;
		xPutSlotCommitted := FALSE;
		xOperationSequenceComplete := FALSE;

